(* IEC 61131-3 sources: daoli-st-library/DL_Process (part 10) *)

(* ---- FC_DL_CathodeMillThroughputCalc.st ---- *)
(*
  Component : FC_DL_CathodeMillThroughputCalc
  Category  : DL_Process
  Function  : 粉碎分级产能估算 t/h：由分级轮转速与风量折算，含转速修正与上限钳位
  Complexity: C2
  开源溯源 : DLF 内部原创（R94 族模板派生）；参考语义来源见 SOURCE_HUNTING_MATRIX.md
  规则遵从 : R1-R16
  契约     : 输入 rAirFlowM3h 系统风量 [m3/h]、rSolidsGm3 气流含尘浓度 [g/m3]、
             nWheelRpm 分级轮实际转速 [r/min]、nWheelRefRpm 分级轮额定转速 [r/min]、
             rSpeedExp 转速修正指数 [-]、rCapMaxTh 产能硬上限 [t/h]；
             输出 rThroughputTh 估算产能 [t/h]、rSpeedFactor 转速修正因子 [-]、
             xCapped 触上限、xValid 有效标志、nFaultCode 故障码。
  边界     : 基础产能 = 风量 × 含尘浓度 / 1.0E6（g→t 与 m3/h→t/h 一次换算）；转速因子 =
             (实际/额定)^指数，指数须 >0 且 ≤2；额定转速为分母须 >1.0E-9 [r/min]；
             产能硬限上限必须具备「极限值→REAL 可表性」反算：上限 1.0E4 [t/h] 远小于 REAL 上限 3.4E38，可表。
  码位     : 9801 输入非有限（故障级）；9802 额定转速或指数越域（故障级）。
*)
FUNCTION FC_DL_CathodeMillThroughputCalc : BOOL
VAR_INPUT
    rAirFlowM3h   : LREAL := 5000.0;   // 系统风量 [m3/h] EN: the air volumetric flow of the classifying system
    rSolidsGm3    : LREAL := 200.0;    // 气流含尘浓度 [g/m3] EN: the solids concentration carried by the air
    nWheelRpm     : INT := 3000;       // 分级轮实际转速 [r/min] EN: the actual rotational speed of the classifying wheel
    nWheelRefRpm  : INT := 3000;       // 分级轮额定转速 [r/min] EN: the rated rotational speed of the classifying wheel
    rSpeedExp     : LREAL := 1.0;      // 转速修正指数 [-] EN: the exponent of the speed correction
    rCapMaxTh     : LREAL := 5.0;      // 产能硬上限 [t/h] EN: the hard upper bound of the throughput
END_VAR
VAR_OUTPUT
    rThroughputTh : LREAL;             // 估算产能 [t/h] EN: the estimated throughput in tonnes per hour
    rSpeedFactor  : LREAL;             // 转速修正因子 [-] EN: the speed correction factor
    xCapped       : BOOL;              // 触产能硬上限 EN: the throughput reached the hard upper bound
    xValid        : BOOL;              // 输出可信标志 EN: the outputs are valid
    nFaultCode    : INT;               // 0=无故障 9801=输入非有限 9802=额定转速或指数越域 EN: zero none, 9801 non finite input, 9802 rated speed or exponent out of range
END_VAR
VAR
    xFinAll : BOOL;                    // 浮点入参同时有限 EN: the floating inputs are finite
    rBase   : LREAL;                   // 基础产能（未修正） [t/h] EN: the base throughput before the correction
    rRatio  : LREAL;                   // 转速比 [-] EN: the speed ratio
    rFactor : LREAL;                   // 修正因子中间值 [-] EN: the interim correction factor
    rOut    : LREAL;                   // 产能中间值 [t/h] EN: the interim throughput
END_VAR
VAR CONSTANT
    DL_CMT_Z       : LREAL := 0.0;      // 浮点零常量 EN: the floating point zero constant
    DL_CMT_MILLION : LREAL := 1.0E6;    // 克转吨与每小时一次换算系数 EN: the gram to tonne conversion factor
    DL_CMT_EXP_MAX : LREAL := 2.0;      // 修正指数上限 [-] EN: the upper bound of the exponent
    DL_CMT_MIN     : LREAL := 1.0E-9;   // 分母绝对值下限 EN: the lower bound of the divisor magnitude
    DL_CMT_C_BAD   : INT := 9801;       // 输入非有限 EN: a non finite input
    DL_CMT_C_RANGE : INT := 9802;       // 额定转速或指数越域 EN: the rated speed or the exponent is out of range
END_VAR

// 段1｜出口预置
FC_DL_CathodeMillThroughputCalc := FALSE;   // 返回值预置假 EN: preset the return value to false
rThroughputTh := DL_CMT_Z;                  // 产能预置零 [t/h] EN: preset the throughput to zero
rSpeedFactor := DL_CMT_Z;                   // 修正因子预置零 [-] EN: preset the correction factor to zero
xCapped := FALSE;                           // 触限标志预置假 EN: preset the capped flag to false
xValid := FALSE;                            // 有效标志预置假 EN: preset the validity flag to false
nFaultCode := 0;                            // 故障码预置零 EN: preset the fault code to zero

// 段2｜非有限闸：浮点入参全列（硬上限参与钳位，漏则钳位失效）
xFinAll := (rAirFlowM3h = rAirFlowM3h) AND ((rAirFlowM3h - rAirFlowM3h) = DL_CMT_Z)
        AND (rSolidsGm3 = rSolidsGm3) AND ((rSolidsGm3 - rSolidsGm3) = DL_CMT_Z)
        AND (rSpeedExp = rSpeedExp) AND ((rSpeedExp - rSpeedExp) = DL_CMT_Z)
        AND (rCapMaxTh = rCapMaxTh) AND ((rCapMaxTh - rCapMaxTh) = DL_CMT_Z);   // 四浮点输入有限性 EN: the finiteness of the four floating inputs
IF NOT xFinAll THEN                                                             // 非有限出口 EN: leave early on a non finite input
    nFaultCode := DL_CMT_C_BAD;                                                 // 非有限码 EN: the non finite code
    RETURN;                                                                     // 早退 EN: return early
END_IF

// 段3｜域闸：风量与含尘浓度非负、转速非负、额定转速过分母下限、指数在 (0,2]、硬上限为正
IF (rAirFlowM3h < DL_CMT_Z) OR (rSolidsGm3 < DL_CMT_Z) OR (nWheelRpm < 0) OR (nWheelRefRpm < 0)
   OR (rSpeedExp <= DL_CMT_Z) OR (rSpeedExp > DL_CMT_EXP_MAX) OR (rCapMaxTh <= DL_CMT_Z)
   OR (ABS(INT_TO_LREAL(nWheelRefRpm)) < DL_CMT_MIN) THEN
    nFaultCode := DL_CMT_C_RANGE;                                               // 越域码 EN: the out of range code
    RETURN;                                                                     // 早退 EN: return early
END_IF

// 段4｜主体：基础产能 = 风量 × 含尘 / 1.0E6；因子 = (实际/额定)^指数
rBase := (rAirFlowM3h * rSolidsGm3) / DL_CMT_MILLION;                           // 基础产能 [t/h] EN: the base throughput
rRatio := INT_TO_LREAL(nWheelRpm) / INT_TO_LREAL(nWheelRefRpm);                 // 转速比，分母已证正 [-] EN: the speed ratio, the divisor is proven positive
rFactor := EXP(rSpeedExp * LN(rRatio));                                         // 指数修正 = e^(k·ln r) [-]，避免依赖 EXPT 方言 EN: the exponential correction without a vendor power operator
rOut := rBase * rFactor;                                                        // 修正后产能 [t/h] EN: the corrected throughput

// 段5｜结果复检 + 硬上限钳位（只防上溢，不下抬）
IF (rOut <> rOut) OR (rOut < DL_CMT_Z) THEN                                     // 复检：非有限或负 EN: recheck for a non finite or negative result
    nFaultCode := DL_CMT_C_RANGE;                                               // 复检失败码 EN: the recheck failure code
    RETURN;                                                                     // 早退，出口保持零哨兵 EN: return early with the zero sentinels
END_IF
IF rOut > rCapMaxTh THEN                                                        // 硬上限钳位 EN: the hard upper bound
    rOut := rCapMaxTh;                                                          // 钳到上限 [t/h] EN: clamp to the upper bound
    xCapped := TRUE;                                                            // 置触限标志 EN: raise the capped flag
END_IF

// 段6｜出口
rThroughputTh := rOut;                                                          // 产能出口 [t/h] EN: the throughput output
rSpeedFactor := rFactor;                                                        // 因子出口 [-] EN: the factor output
xValid := TRUE;                                                                 // 结果可信 EN: the results are valid
FC_DL_CathodeMillThroughputCalc := TRUE;                                        // 返回真 EN: return true
END_FUNCTION

(* ---- FC_DL_CathodeMoistureSpecCalc.st ---- *)
(*
  Component : FC_DL_CathodeMoistureSpecCalc
  Category  : DL_Process
  Function  : 水分限值与所需干燥时间反算（一阶指数干燥模型 t = -τ × LN(M目标/M初始)）
  Complexity: C2
  开源溯源 : DLF 内部原创（R94 族模板派生）；参考语义来源见 SOURCE_HUNTING_MATRIX.md
  规则遵从 : R1-R16
  契约     : 输入 rMoistInitPct 初始水分 [%]、rMoistTargetPct 目标水分限值 [%]、
             rDryTauMin 干燥时间常数 [min]、rDryTimeMaxMin 工艺允许最长干燥时间 [min]；
             输出 rDryMin 计算所需干燥时间 [min]、rMoistRatio 水分比 [-]、
             xSpecAchievable 目标在当前允许时间内可达、xValid 有效标志、nFaultCode 故障码。
  边界     : 须 初始水分 > 目标水分 > 0；时间常数为分母须 >1.0E-9 [min]；允许时长须 >0；
             模型不含恒速段与临界含水率，仅适用于降速干燥段（物料表面已不饱和）；
             目标不可达只置 xSpecAchievable=FALSE 为信息级，不置故障。
  码位     : 9801 输入非有限（故障级）；9802 水分关系非法（故障级）；9803 时间常数或允许时长越域（故障级）。
*)
FUNCTION FC_DL_CathodeMoistureSpecCalc : BOOL
VAR_INPUT
    rMoistInitPct   : LREAL := 5.0;      // 初始水分 [%] EN: the initial moisture content
    rMoistTargetPct : LREAL := 0.05;     // 目标水分限值 [%] EN: the target moisture limit
    rDryTauMin      : LREAL := 20.0;     // 干燥时间常数 [min] EN: the drying time constant
    rDryTimeMaxMin  : LREAL := 180.0;    // 工艺允许最长干燥时间 [min] EN: the longest drying time allowed by the process
END_VAR
VAR_OUTPUT
    rDryMin         : LREAL;             // 计算所需干燥时间 [min] EN: the computed drying time required
    rMoistRatio     : LREAL;             // 目标与初始水分之比 [-] EN: the ratio of the target to the initial moisture
    xSpecAchievable : BOOL;              // 目标在允许时间内可达（信息级） EN: the target is reachable within the allowed time, information class only
    xValid          : BOOL;              // 输出可信标志 EN: the outputs are valid
    nFaultCode      : INT;               // 0=无故障 9801=输入非有限 9802=水分关系非法 9803=常数或时长越域 EN: zero none, 9801 non finite, 9802 illegal moisture relation, 9803 constant or duration out of range
END_VAR
VAR
    xFinAll : BOOL;                      // 四输入同时有限 EN: all four inputs are finite
    rRat    : LREAL;                     // 水分比中间值 [-] EN: the interim moisture ratio
    rLn     : LREAL;                     // 水分比对数 [-] EN: the logarithm of the moisture ratio
    rT      : LREAL;                     // 干燥时间中间值 [min] EN: the interim drying time
END_VAR
VAR CONSTANT
    DL_CMS_Z      : LREAL := 0.0;        // 浮点零常量 EN: the floating point zero constant
    DL_CMS_MIN    : LREAL := 1.0E-9;     // 分母绝对值下限 EN: the lower bound of the divisor magnitude
    DL_CMS_C_BAD  : INT := 9801;         // 输入非有限 EN: a non finite input
    DL_CMS_C_REL  : INT := 9802;         // 水分关系非法 EN: an illegal moisture relation
    DL_CMS_C_RANG : INT := 9803;         // 时间常数或允许时长越域 EN: the constant or the duration is out of range
END_VAR

// 段1｜出口预置
FC_DL_CathodeMoistureSpecCalc := FALSE;   // 返回值预置假 EN: preset the return value to false
rDryMin := DL_CMS_Z;                      // 干燥时间预置零 [min] EN: preset the drying time to zero
rMoistRatio := DL_CMS_Z;                  // 水分比预置零 [-] EN: preset the moisture ratio to zero
xSpecAchievable := FALSE;                 // 可达标志预置假 EN: preset the reachability flag to false
xValid := FALSE;                          // 有效标志预置假 EN: preset the validity flag to false
nFaultCode := 0;                          // 故障码预置零 EN: preset the fault code to zero

// 段2｜非有限闸：四输入全列
xFinAll := (rMoistInitPct = rMoistInitPct) AND ((rMoistInitPct - rMoistInitPct) = DL_CMS_Z)
        AND (rMoistTargetPct = rMoistTargetPct) AND ((rMoistTargetPct - rMoistTargetPct) = DL_CMS_Z)
        AND (rDryTauMin = rDryTauMin) AND ((rDryTauMin - rDryTauMin) = DL_CMS_Z)
        AND (rDryTimeMaxMin = rDryTimeMaxMin) AND ((rDryTimeMaxMin - rDryTimeMaxMin) = DL_CMS_Z);   // 四输入有限性 EN: the finiteness of all four inputs
IF NOT xFinAll THEN                                                                                 // 非有限出口 EN: leave early on a non finite input
    nFaultCode := DL_CMS_C_BAD;                                                                     // 非有限码 EN: the non finite code
    RETURN;                                                                                         // 早退 EN: return early
END_IF

// 段3｜域闸：水分关系 初始 > 目标 > 0；时间常数与允许时长为正
IF (rMoistTargetPct <= DL_CMS_Z) OR (rMoistInitPct <= rMoistTargetPct) THEN                          // 水分关系闸 EN: the moisture relation gate
    nFaultCode := DL_CMS_C_REL;                                                                     // 关系非法码 EN: the relation code
    RETURN;                                                                                         // 早退 EN: return early
END_IF
IF (rDryTauMin < DL_CMS_MIN) OR (rDryTimeMaxMin <= DL_CMS_Z) THEN                                    // 常数与时长闸 EN: the constant and duration gate
    nFaultCode := DL_CMS_C_RANG;                                                                    // 越域码 EN: the out of range code
    RETURN;                                                                                         // 早退 EN: return early
END_IF

// 段4｜主体：t = -τ × LN(目标/初始)，比值已证在 (0,1)
rRat := rMoistTargetPct / rMoistInitPct;                                                            // 水分比 [-] EN: the moisture ratio
rLn := LN(rRat);                                                                                    // 水分比对数，已证 <0 [-] EN: the logarithm of the ratio, proven negative
rT := -rDryTauMin * rLn;                                                                            // 所需干燥时间 [min] EN: the drying time required
IF (rT <> rT) OR (rT < DL_CMS_Z) THEN                                                               // 结果复检 EN: recheck the result
    nFaultCode := DL_CMS_C_RANG;                                                                    // 复检失败码 EN: the recheck failure code
    RETURN;                                                                                         // 早退，出口保持零哨兵 EN: return early with the zero sentinels
END_IF

// 段5｜出口：可达性为信息级判据
rDryMin := rT;                                                                                      // 干燥时间出口 [min] EN: the drying time output
rMoistRatio := rRat;                                                                                // 水分比出口 [-] EN: the moisture ratio output
xSpecAchievable := rT <= rDryTimeMaxMin;                                                            // 可达性判定 EN: the reachability verdict
xValid := TRUE;                                                                                     // 结果可信 EN: the results are valid
FC_DL_CathodeMoistureSpecCalc := TRUE;                                                              // 返回真 EN: return true
END_FUNCTION

(* ---- FC_DL_CathodeO2PartialPressureCalc.st ---- *)
(*
  Component : FC_DL_CathodeO2PartialPressureCalc
  Category  : DL_Process
  Function  : 烧结气氛氧分压 = 氧体积浓度 × 总压，并统一换算到 kPa
  Complexity: C2
  开源溯源 : DLF 内部原创（R94 族模板派生）；参考语义来源见 SOURCE_HUNTING_MATRIX.md
  规则遵从 : R1-R16
  契约     : 输入 rO2Pct 氧体积浓度 [%]、rTotalPressKpa 炉膛总压 [kPa]、rO2LowKpa 氧分压下限 [kPa]；
             输出 rPO2Kpa 氧分压 [kPa]、rO2Ppm 氧体积浓度折算 [ppm]、xO2Low 低于下限（信息级）、
             xValid 有效标志、nFaultCode 故障码。
  边界     : 氧浓度须在 0~100 [%] 内、总压须 >std 0（表压与绝压口径由调用方统一为绝压）；
             浓度 1 [%] = 10000 [ppm]，故 ppm = % × 10000；本件为绝压口径，不做大气压叠加。
  码位     : 9801 输入非有限（故障级）；9802 浓度或总压越域（故障级）。
*)
FUNCTION FC_DL_CathodeO2PartialPressureCalc : BOOL
VAR_INPUT
    rO2Pct       : LREAL := 21.0;     // 氧体积浓度 [%] EN: the oxygen volumetric concentration in percent
    rTotalPressKpa: LREAL := 101.325; // 炉膛总压（绝压口径） [kPa] EN: the furnace total pressure on the absolute scale
    rO2LowKpa    : LREAL := 0.5;      // 氧分压工艺下限 [kPa] EN: the technological lower bound of the oxygen partial pressure
END_VAR
VAR_OUTPUT
    rPO2Kpa : LREAL;                  // 氧分压 [kPa] EN: the oxygen partial pressure
    rO2Ppm  : LREAL;                  // 氧体积浓度折算值 [ppm] EN: the oxygen concentration expressed in ppm
    xO2Low  : BOOL;                   // 氧分压低于工艺下限（信息级） EN: the oxygen partial pressure is below the limit, information class only
    xValid  : BOOL;                   // 输出可信标志 EN: the outputs are valid
    nFaultCode : INT;                 // 0=无故障 9801=输入非有限 9802=浓度或总压越域 EN: zero none, 9801 non finite input, 9802 concentration or pressure out of range
END_VAR
VAR
    xFinAll : BOOL;                   // 三输入同时有限 EN: all three inputs are finite
    rFrac   : LREAL;                  // 氧体积分数 [-] EN: the oxygen volumetric fraction
    rPO2    : LREAL;                  // 氧分压中间值 [kPa] EN: the interim oxygen partial pressure
    rPpm    : LREAL;                  // ppm 中间值 [ppm] EN: the interim ppm value
END_VAR
VAR CONSTANT
    DL_COP_Z         : LREAL := 0.0;      // 浮点零常量 EN: the floating point zero constant
    DL_COP_HUNDRED   : LREAL := 100.0;    // 百分数换算系数 EN: the percent conversion factor
    DL_COP_PPM_FACT  : LREAL := 10000.0;  // 百分数转 ppm 的系数 EN: the percent to ppm factor
    DL_COP_C_BAD     : INT := 9801;       // 输入非有限 EN: a non finite input
    DL_COP_C_RANGE   : INT := 9802;       // 浓度或总压越域 EN: the concentration or the pressure is out of range
END_VAR

// 段1｜出口预置
FC_DL_CathodeO2PartialPressureCalc := FALSE;   // 返回值预置假 EN: preset the return value to false
rPO2Kpa := DL_COP_Z;                           // 氧分压预置零 [kPa] EN: preset the partial pressure to zero
rO2Ppm := DL_COP_Z;                            // ppm 预置零 [ppm] EN: preset the ppm value to zero
xO2Low := FALSE;                               // 低压标志预置假 EN: preset the low pressure flag to false
xValid := FALSE;                               // 有效标志预置假 EN: preset the validity flag to false
nFaultCode := 0;                               // 故障码预置零 EN: preset the fault code to zero

// 段2｜非有限闸：三输入全列（下限参与出口判据）
xFinAll := (rO2Pct = rO2Pct) AND ((rO2Pct - rO2Pct) = DL_COP_Z)
        AND (rTotalPressKpa = rTotalPressKpa) AND ((rTotalPressKpa - rTotalPressKpa) = DL_COP_Z)
        AND (rO2LowKpa = rO2LowKpa) AND ((rO2LowKpa - rO2LowKpa) = DL_COP_Z);   // 三输入有限性 EN: the finiteness of all three inputs
IF NOT xFinAll THEN                                                             // 非有限出口 EN: leave early on a non finite input
    nFaultCode := DL_COP_C_BAD;                                                 // 输入非有限码 EN: the non finite code
    RETURN;                                                                     // 早退 EN: return early
END_IF

// 段3｜域闸：氧浓度 0~100 [%]、总压为正、下限非负
IF (rO2Pct < DL_COP_Z) OR (rO2Pct > DL_COP_HUNDRED) OR (rTotalPressKpa <= DL_COP_Z)
   OR (rO2LowKpa < DL_COP_Z) THEN
    nFaultCode := DL_COP_C_RANGE;                                               // 越域码 EN: the out of range code
    RETURN;                                                                     // 早退 EN: return early
END_IF

// 段4｜主体：pO2 = 浓度/100 × 总压；ppm = 浓度 × 10000
rFrac := rO2Pct / DL_COP_HUNDRED;                                               // 氧体积分数 [-] EN: the oxygen volumetric fraction
rPO2 := rFrac * rTotalPressKpa;                                                 // 氧分压 [kPa] EN: the oxygen partial pressure
rPpm := rO2Pct * DL_COP_PPM_FACT;                                               // 浓度转 ppm [ppm] EN: the concentration in ppm

// 段5｜出口
rPO2Kpa := rPO2;                                                                // 氧分压出口 [kPa] EN: the partial pressure output
rO2Ppm := rPpm;                                                                 // ppm 出口 [ppm] EN: the ppm output
xO2Low := rPO2 < rO2LowKpa;                                                     // 低压判据（信息级） EN: the low pressure test, information class only
xValid := TRUE;                                                                 // 结果可信 EN: the results are valid
FC_DL_CathodeO2PartialPressureCalc := TRUE;                                     // 返回真 EN: return true
END_FUNCTION

(* ---- FC_DL_CathodeSaggerLoadCalc.st ---- *)
(*
  Component : FC_DL_CathodeSaggerLoadCalc
  Category  : DL_Process
  Function  : 匣钵装载量 = 层数 × 每层片数 × 单重，并做超重告警
  Complexity: C2
  开源溯源 : DLF 内部原创（R94 族模板派生）；参考语义来源见 SOURCE_HUNTING_MATRIX.md
  规则遵从 : R1-R16
  契约     : 输入 nLayers 层数 [层]、nPerLayer 每层片数 [片/层]、rPieceKg 单片重量 [kg]、
             rMaxLoadKg 匣钵允许装载上限 [kg]；输出 nPieceCount 总片数 [片]、rLoadKg 装载总重 [kg]、
             xOverload 超重（故障级：超重会导致匣钵破裂并损坏辊棒，按安全侧立即判故障）、
             xValid 有效标志、nFaultCode 故障码。
  边界     : 层数与每层片数须在 0~999 内（超过 999 属组态错误，防整数乘法溢出判 9802）；
             单片重量须 ≥0；上限须 >0；总片数 = 层数 × 每层片数，最大 999×999 = 998001 片，INT 可表；
             超重按方向明确判「超上限」，故为故障级（R146：与安全侧一致的异常立即终止）。
  码位     : 9801 输入非有限或为负（故障级）；9802 计数越界（故障级）；9803 超重（故障级）。
*)
FUNCTION FC_DL_CathodeSaggerLoadCalc : BOOL
VAR_INPUT
    nLayers    : INT := 8;           // 匣钵叠放层数 [层] EN: the number of stacked layers in the sagger
    nPerLayer  : INT := 6;           // 每层片数 [片/层] EN: the number of pieces per layer
    rPieceKg   : LREAL := 0.5;       // 单片重量 [kg] EN: the weight of one piece
    rMaxLoadKg : LREAL := 30.0;      // 匣钵允许装载上限 [kg] EN: the allowed load limit of the sagger
END_VAR
VAR_OUTPUT
    nPieceCount : INT;               // 总片数 [片] EN: the total piece count
    rLoadKg     : LREAL;             // 装载总重 [kg] EN: the total load weight
    xOverload   : BOOL;              // 超重（故障级） EN: the load exceeds the limit, a fault class condition
    xValid      : BOOL;              // 输出可信标志 EN: the outputs are valid
    nFaultCode  : INT;               // 0=无故障 9801=输入非法 9802=计数越界 9803=超重 EN: zero none, 9801 illegal input, 9802 count out of range, 9803 overload
END_VAR
VAR
    xFinAll  : BOOL;                 // 两个浮点入参有限 EN: both floating inputs are finite
    nCnt     : INT;                  // 总片数中间值 [片] EN: the interim piece count
    rLoad    : LREAL;                // 总重中间值 [kg] EN: the interim load weight
END_VAR
VAR CONSTANT
    DL_CSL_Z      : LREAL := 0.0;    // 浮点零常量 EN: the floating point zero constant
    DL_CSL_CNT_MAX: INT := 999;      // 层数与每层片数上限 [个] EN: the upper bound of the layer count and the per layer count
    DL_CSL_C_BAD  : INT := 9801;     // 输入非法 EN: an illegal input
    DL_CSL_C_CNT  : INT := 9802;     // 计数越界 EN: the count is out of range
    DL_CSL_C_OVER : INT := 9803;     // 超重 EN: the overload condition
END_VAR

// 段1｜出口预置
FC_DL_CathodeSaggerLoadCalc := FALSE;   // 返回值预置假 EN: preset the return value to false
nPieceCount := 0;                        // 总片数预置零 [片] EN: preset the piece count to zero
rLoadKg := DL_CSL_Z;                     // 总重预置零 [kg] EN: preset the load weight to zero
xOverload := FALSE;                      // 超重标志预置假 EN: preset the overload flag to false
xValid := FALSE;                         // 有效标志预置假 EN: preset the validity flag to false
nFaultCode := 0;                         // 故障码预置零 EN: preset the fault code to zero

// 段2｜非有限闸：两个浮点入参全列（上限参与超重判据）
xFinAll := (rPieceKg = rPieceKg) AND ((rPieceKg - rPieceKg) = DL_CSL_Z)
        AND (rMaxLoadKg = rMaxLoadKg) AND ((rMaxLoadKg - rMaxLoadKg) = DL_CSL_Z);   // 两输入有限性 EN: the finiteness of both inputs
IF NOT xFinAll THEN                                                                 // 非有限出口 EN: leave early on a non finite input
    nFaultCode := DL_CSL_C_BAD;                                                     // 输入非法码 EN: the illegal input code
    RETURN;                                                                         // 早退 EN: return early
END_IF

// 段3｜域闸：单片重量与上限为正、两计数非负且不超 999
IF (rPieceKg < DL_CSL_Z) OR (rMaxLoadKg <= DL_CSL_Z) THEN                            // 数值域闸 EN: the numeric domain gate
    nFaultCode := DL_CSL_C_BAD;                                                     // 输入非法码 EN: the illegal input code
    RETURN;                                                                         // 早退 EN: return early
END_IF
IF (nLayers < 0) OR (nLayers > DL_CSL_CNT_MAX) OR (nPerLayer < 0) OR (nPerLayer > DL_CSL_CNT_MAX) THEN
    nFaultCode := DL_CSL_C_CNT;                                                     // 计数越界码 EN: the count out of range code
    RETURN;                                                                         // 早退 EN: return early
END_IF

// 段4｜主体：片数用整数乘（取值范围已证），重量用标准转换后相乘
nCnt := nLayers * nPerLayer;                                                        // 总片数 [片] EN: the total piece count
rLoad := INT_TO_LREAL(nCnt) * rPieceKg;                                             // 总重 [kg] EN: the total load weight

// 段5｜出口：超重为故障级（安全侧一致的方向明确异常立即终止）
nPieceCount := nCnt;                                                                // 总片数出口 [片] EN: the piece count output
rLoadKg := rLoad;                                                                   // 总重出口 [kg] EN: the load weight output
IF rLoad > rMaxLoadKg THEN                                                          // 超重判据 EN: the overload test
    xOverload := TRUE;                                                              // 置超重标志 EN: raise the overload flag
    nFaultCode := DL_CSL_C_OVER;                                                    // 超重码 EN: the overload code
    xValid := FALSE;                                                                // 超重时输出不可用于投料 EN: the outputs are not usable for loading
    RETURN;                                                                         // 早退（返回假） EN: return false
END_IF
xValid := TRUE;                                                                     // 结果可信 EN: the results are valid
FC_DL_CathodeSaggerLoadCalc := TRUE;                                                // 返回真 EN: return true
END_FUNCTION

(* ---- FC_DL_CathodeSinterSoakCalc.st ---- *)
(*
  Component : FC_DL_CathodeSinterSoakCalc
  Category  : DL_Process
  Function  : 烧结保温时间由固相扩散长度与粒径反算，t = L² / (4D)，含最小值保护
  Complexity: C2
  开源溯源 : DLF 内部原创（R94 族模板派生）；参考语义来源见 SOURCE_HUNTING_MATRIX.md
  规则遵从 : R1-R16
  契约     : 输入 rDiffLenUm 目标扩散长度 [μm]、rDiffCoefUm2Min 有效扩散系数 [μm2/min]、
             rParticleD50Um 一次粒径中位径 [μm]、rSoakMinMin 保温时间下限 [min]；
             输出 rSoakCalcMin 模型计算保温时间 [min]、rSoakMin 施加下限保护后的保温时间 [min]、
             xMinApplied 触底保护生效、xValid 有效标志、nFaultCode 故障码。
  边界     : 扩散系数为分母须 >1.0E-9 [μm2/min]；扩散长度与粒径须 >0；模型 t = L²/(4D)；
             粒径小于两倍扩散长度时扩散已贯穿颗粒，模型外推无意义，rSoakMin 仍给出但不置 xValid=FALSE，
             改由 xMinApplied 与告警表达（本件不设粒径下限门限，交由上层工艺判定）。
  码位     : 9801 输入非法（故障级）；9802 扩散系数过小（故障级）。
*)
FUNCTION FC_DL_CathodeSinterSoakCalc : BOOL
VAR_INPUT
    rDiffLenUm      : LREAL := 2.0;      // 目标固相扩散长度 [μm] EN: the target solid state diffusion length
    rDiffCoefUm2Min : LREAL := 0.05;     // 有效扩散系数 [μm2/min] EN: the effective diffusion coefficient
    rParticleD50Um  : LREAL := 5.0;      // 一次粒径中位径 D50 [μm] EN: the median primary particle size
    rSoakMinMin     : LREAL := 120.0;    // 保温时间工艺下限 [min] EN: the technological lower bound of the soak time
END_VAR
VAR_OUTPUT
    rSoakCalcMin : LREAL;                // 模型计算保温时间 [min] EN: the model computed soak time
    rSoakMin     : LREAL;                // 施加下限保护后的保温时间 [min] EN: the soak time after the lower bound protection
    xMinApplied  : BOOL;                 // 触底保护生效 EN: the lower bound protection took effect
    xThrough     : BOOL;                 // 扩散已贯穿颗粒（信息级） EN: the diffusion length already spans the particle, information class only
    xValid       : BOOL;                 // 输出可信标志 EN: the outputs are valid
    nFaultCode   : INT;                  // 0=无故障 9801=输入非法 9802=扩散系数过小 EN: zero none, 9801 illegal input, 9802 diffusion coefficient too small
END_VAR
VAR
    xFinAll  : BOOL;                     // 四输入同时有限 EN: all four inputs are finite
    rDen     : LREAL;                    // 分母 4D [μm2/min] EN: the divisor, four times the diffusion coefficient
    rSq      : LREAL;                    // 扩散长度平方 [μm2] EN: the squared diffusion length
    rCalc    : LREAL;                    // 计算保温时间 [min] EN: the computed soak time
    rApply   : LREAL;                    // 施加下限后的保温时间 [min] EN: the soak time after the lower bound
END_VAR
VAR CONSTANT
    DL_CSS_Z       : LREAL := 0.0;       // 浮点零常量 EN: the floating point zero constant
    DL_CSS_FOUR    : LREAL := 4.0;       // 扩散方程几何系数 EN: the geometric factor of the diffusion equation
    DL_CSS_TWO     : LREAL := 2.0;       // 贯穿判据倍数 EN: the spanning criterion multiplier
    DL_CSS_MIN     : LREAL := 1.0E-9;    // 分母绝对值下限 [μm2/min] EN: the lower bound of the divisor magnitude
    DL_CSS_C_BAD   : INT := 9801;        // 输入非法 EN: an illegal input
    DL_CSS_C_COEF  : INT := 9802;        // 扩散系数过小 EN: the diffusion coefficient is too small
END_VAR

// 段1｜出口预置
FC_DL_CathodeSinterSoakCalc := FALSE;   // 返回值预置假 EN: preset the return value to false
rSoakCalcMin := DL_CSS_Z;               // 计算保温时间预置零 [min] EN: preset the computed soak time to zero
rSoakMin := DL_CSS_Z;                   // 施加下限后保温时间预置零 [min] EN: preset the final soak time to zero
xMinApplied := FALSE;                   // 触底标志预置假 EN: preset the lower bound flag to false
xThrough := FALSE;                      // 贯穿标志预置假 EN: preset the spanning flag to false
xValid := FALSE;                        // 有效标志预置假 EN: preset the validity flag to false
nFaultCode := 0;                        // 故障码预置零 EN: preset the fault code to zero

// 段2｜非有限闸：四输入全列
xFinAll := (rDiffLenUm = rDiffLenUm) AND ((rDiffLenUm - rDiffLenUm) = DL_CSS_Z)
        AND (rDiffCoefUm2Min = rDiffCoefUm2Min) AND ((rDiffCoefUm2Min - rDiffCoefUm2Min) = DL_CSS_Z)
        AND (rParticleD50Um = rParticleD50Um) AND ((rParticleD50Um - rParticleD50Um) = DL_CSS_Z)
        AND (rSoakMinMin = rSoakMinMin) AND ((rSoakMinMin - rSoakMinMin) = DL_CSS_Z);   // 四输入有限性 EN: the finiteness of all four inputs
IF NOT xFinAll THEN                                                                      // 非有限出口 EN: leave early on a non finite input
    nFaultCode := DL_CSS_C_BAD;                                                          // 输入非法码 EN: the illegal input code
    RETURN;                                                                              // 早退 EN: return early
END_IF

// 段3｜域闸：扩散长度、粒径为正；扩散系数过分母下限；下限时间非负
rDen := DL_CSS_FOUR * rDiffCoefUm2Min;                                                   // 分母 4D [μm2/min] EN: the divisor, four times the diffusion coefficient
IF (rDiffLenUm <= DL_CSS_Z) OR (rParticleD50Um <= DL_CSS_Z) OR (rSoakMinMin < DL_CSS_Z)
   OR (ABS(rDen) < DL_CSS_MIN) THEN
    nFaultCode := DL_CSS_C_COEF;                                                         // 系数或域非法码 EN: the coefficient or domain code
    RETURN;                                                                              // 早退 EN: return early
END_IF

// 段4｜主体：t = L² / (4D)
rSq := rDiffLenUm * rDiffLenUm;                                                          // 扩散长度平方 [μm2] EN: the squared diffusion length
rCalc := rSq / rDen;                                                                     // 计算保温时间 [min] EN: the computed soak time
IF (rCalc <> rCalc) OR (rCalc < DL_CSS_Z) THEN                                           // 结果复检 EN: recheck the result
    nFaultCode := DL_CSS_C_COEF;                                                         // 复检失败码 EN: the recheck failure code
    RETURN;                                                                              // 早退，出口保持零哨兵 EN: return early with the zero sentinels
END_IF

// 段5｜最小值保护与贯穿标记
rApply := rCalc;                                                                         // 施加下限工作副本 [min] EN: the working copy for the lower bound
xMinApplied := rCalc < rSoakMinMin;                                                      // 触底判据 EN: the lower bound test
IF xMinApplied THEN                                                                      // 触底则抬到工艺下限 EN: raise to the process lower bound
    rApply := rSoakMinMin;                                                               // 施加下限 [min] EN: apply the lower bound
END_IF
xThrough := rDiffLenUm >= (rParticleD50Um / DL_CSS_TWO);                                 // 贯穿判据（信息级） EN: the spanning test, information class only

// 段6｜出口
rSoakCalcMin := rCalc;                                                                   // 计算值出口 [min] EN: the computed value output
rSoakMin := rApply;                                                                      // 最终值出口 [min] EN: the final value output
xValid := TRUE;                                                                          // 结果可信 EN: the results are valid
FC_DL_CathodeSinterSoakCalc := TRUE;                                                     // 返回真 EN: return true
END_FUNCTION

(* ---- FC_DL_CathodeTapDensityCalc.st ---- *)
(*
  Component : FC_DL_CathodeTapDensityCalc
  Category  : DL_Process
  Function  : 振实密度 = 质量 / 振实后体积，并按振次做修正
  Complexity: C2
  开源溯源 : DLF 内部原创（R94 族模板派生）；参考语义来源见 SOURCE_HUNTING_MATRIX.md
  规则遵从 : R1-R16
  契约     : 输入 rMassG 试样质量 [g]、rVolumeMl 振实后体积 [ml]、nTaps 实测振次 [次]、
             nRefTaps 标准振次 [次]、rTapCoef 振次修正系数 [-]；
             输出 rDensityGml 实测振实密度 [g/ml]、rDensityCorrGml 修正到标准振次的密度 [g/ml]、
             xValid 有效标志、nFaultCode 故障码。
  边界     : 体积为分母须 >1.0E-9 [ml]；振次须 ≥1（取对数的前提），标准振次须 ≥1；
             修正模型 rho_ref = rho × (1 + k × LN(nRef/nTaps))，k 须在 [0, 0.2] 内，
             越域判 9803（k 越域会把修正放大成伪数据）；1 g/ml = 1 g/cm3，单位不做换算。
  码位     : 9801 输入非法（故障级）；9802 体积过小或振次非法（故障级）；9803 修正系数越域（故障级）。
*)
FUNCTION FC_DL_CathodeTapDensityCalc : BOOL
VAR_INPUT
    rMassG    : LREAL := 100.0;    // 试样质量 [g] EN: the mass of the sample
    rVolumeMl : LREAL := 50.0;     // 振实后体积 [ml] EN: the tapped volume of the sample
    nTaps     : INT := 3000;       // 实测振次 [次] EN: the tap count actually applied
    nRefTaps  : INT := 3000;       // 标准振次 [次] EN: the reference tap count
    rTapCoef  : LREAL := 0.02;     // 振次修正系数 [-] EN: the tap count correction coefficient
END_VAR
VAR_OUTPUT
    rDensityGml     : LREAL;       // 实测振实密度 [g/ml] EN: the measured tap density
    rDensityCorrGml : LREAL;       // 修正到标准振次的密度 [g/ml] EN: the density corrected to the reference tap count
    xValid          : BOOL;        // 输出可信标志 EN: the outputs are valid
    nFaultCode      : INT;         // 0=无故障 9801=输入非法 9802=体积或振次非法 9803=系数越域 EN: zero none, 9801 illegal input, 9802 volume or taps illegal, 9803 coefficient out of range
END_VAR
VAR
    xFinAll : BOOL;                // 三个浮点入参有限 EN: the three floating inputs are finite
    rDen    : LREAL;               // 分母（振实后体积） [ml] EN: the divisor, the tapped volume
    rRho    : LREAL;               // 实测密度 [g/ml] EN: the measured density
    rLnCorr : LREAL;               // 振次比对数 [-] EN: the logarithm of the tap ratio
    rCorr   : LREAL;               // 密度修正中间值 [g/ml] EN: the interim corrected density
END_VAR
VAR CONSTANT
    DL_CTD_Z        : LREAL := 0.0;   // 浮点零常量 EN: the floating point zero constant
    DL_CTD_ONE      : LREAL := 1.0;   // 浮点壹常量 EN: the floating point one constant
    DL_CTD_COEF_MAX : LREAL := 0.2;   // 修正系数上限 [-] EN: the upper bound of the correction coefficient
    DL_CTD_MIN      : LREAL := 1.0E-9;// 分母绝对值下限 [ml] EN: the lower bound of the divisor magnitude
    DL_CTD_C_BAD    : INT := 9801;    // 输入非法 EN: an illegal input
    DL_CTD_C_DEN    : INT := 9802;    // 体积过小或振次非法 EN: the volume is too small or the taps are illegal
    DL_CTD_C_COEF   : INT := 9803;    // 修正系数越域 EN: the coefficient is out of range
END_VAR

// 段1｜出口预置
FC_DL_CathodeTapDensityCalc := FALSE;   // 返回值预置假 EN: preset the return value to false
rDensityGml := DL_CTD_Z;                 // 实测密度预置零 [g/ml] EN: preset the measured density to zero
rDensityCorrGml := DL_CTD_Z;             // 修正密度预置零 [g/ml] EN: preset the corrected density to zero
xValid := FALSE;                         // 有效标志预置假 EN: preset the validity flag to false
nFaultCode := 0;                         // 故障码预置零 EN: preset the fault code to zero

// 段2｜非有限闸：三浮点入参全列
xFinAll := (rMassG = rMassG) AND ((rMassG - rMassG) = DL_CTD_Z)
        AND (rVolumeMl = rVolumeMl) AND ((rVolumeMl - rVolumeMl) = DL_CTD_Z)
        AND (rTapCoef = rTapCoef) AND ((rTapCoef - rTapCoef) = DL_CTD_Z);   // 三输入有限性 EN: the finiteness of all three inputs
IF NOT xFinAll THEN                                                        // 非有限出口 EN: leave early on a non finite input
    nFaultCode := DL_CTD_C_BAD;                                            // 输入非法码 EN: the illegal input code
    RETURN;                                                                // 早退 EN: return early
END_IF

// 段3｜域闸：质量为非负、体积过分母下限、振次 ≥1
rDen := rVolumeMl;                                                          // 取分母 [ml] EN: take the divisor
IF (rMassG < DL_CTD_Z) OR (ABS(rDen) < DL_CTD_MIN) OR (nTaps < 1) OR (nRefTaps < 1) THEN
    nFaultCode := DL_CTD_C_DEN;                                            // 体积或振次非法码 EN: the volume or tap code
    RETURN;                                                                // 早退 EN: return early
END_IF
IF (rTapCoef < DL_CTD_Z) OR (rTapCoef > DL_CTD_COEF_MAX) THEN               // 系数域闸 EN: the coefficient domain gate
    nFaultCode := DL_CTD_C_COEF;                                            // 系数越域码 EN: the coefficient code
    RETURN;                                                                // 早退 EN: return early
END_IF

// 段4｜主体：实测密度与振次修正（两出口同源，修正只缩放实测值不另起公式）
rRho := rMassG / rDen;                                                      // 实测振实密度 [g/ml] EN: the measured tap density
rLnCorr := LN(INT_TO_LREAL(nRefTaps) / INT_TO_LREAL(nTaps));                // 振次比对数 [-]，两者已证 ≥1 EN: the logarithm of the tap ratio
rCorr := rRho * (DL_CTD_ONE + rTapCoef * rLnCorr);                          // 修正密度 [g/ml] EN: the corrected density
IF (rCorr <> rCorr) OR (rCorr < DL_CTD_Z) THEN                              // 结果复检 EN: recheck the result
    nFaultCode := DL_CTD_C_COEF;                                            // 复检失败码 EN: the recheck failure code
    rDensityGml := rRho;                                                    // 实测值仍可给出 EN: the measured value is still published
    RETURN;                                                                // 早退 EN: return early
END_IF

// 段5｜出口
rDensityGml := rRho;                                                        // 实测密度出口 [g/ml] EN: the measured density output
rDensityCorrGml := rCorr;                                                   // 修正密度出口 [g/ml] EN: the corrected density output
xValid := TRUE;                                                             // 结果可信 EN: the results are valid
FC_DL_CathodeTapDensityCalc := TRUE;                                        // 返回真 EN: return true
END_FUNCTION

(* ---- FC_DL_CellOccupyRateCalc.st ---- *)
(*
  ============================================================
  组件名 : FC_DL_CellOccupyRateCalc
  分类   : DL_Process
  功能   : 货位占用率计算，扣除封存货位后按可用货位求占用百分比与空闲数
  复杂度 : C1
  版本   : 1.0.0
  作者   : 道莅工业代码库工厂 / R81
  日期   : 2026-11-24
  开源溯源 : clean-room（no upstream）—— 依据公开工程公式自研，未复制任何上游实现
  红线自检 : R1 无GVL/R2 无物理地址/R3 纯IEC/R4 防除零/R5 双语注释
  接口说明 :
      可用货位 = 总货位 - 封存货位；占用率 = 已用 / 可用 * 100。
      可用货位 <= 0 时占用率无定义，直接判无效，不输出替代值。
      空闲货位 = 可用 - 已用，小于 0 表示超占（数据异常），本实现按 0 截断并保持比例可算。
      中间量用 DINT 承载，避免 INT 减法溢出。
  ============================================================
*)
FUNCTION FC_DL_CellOccupyRateCalc : BOOL
VAR_INPUT
    bEnable       : BOOL; // 使能：TRUE 时计算 / Enable: TRUE to compute
    bErr          : BOOL; // 外部故障：TRUE 时立即退出并置结果无效 / External fault: TRUE aborts with invalid result
    iCellTotal    : INT;  // 货位总数量 [个] / total number of storage cells [unit]
    iCellUsed     : INT;  // 已占用货位数量 [个] / number of occupied cells [unit]
    iCellBlocked  : INT;  // 封存禁用货位数量 [个] / number of blocked or disabled cells [unit]
END_VAR
VAR_OUTPUT
    rOccupyPct : REAL; // 可用货位占用率 [%] / occupancy rate over the available cells [percent]
    iCellFree  : INT;  // 空闲货位数量，负值按 0 截断 [个] / free cell count, negative clamped to zero [unit]
    iCellAvail : INT;  // 扣除封存后的可用货位数量 [个] / available cell count after removing blocked cells [unit]
    bValid     : BOOL; // 输出有效：TRUE 表示结果可用 / Output valid
END_VAR
VAR CONSTANT
    DL_R_MAX : REAL := 3.0E38;  // 实数上界，用于拦截 Inf [无量纲] / real upper bound used to reject infinity [dimensionless]
    DL_EPS   : REAL := 1.0E-12; // 除零判定阈值 [无量纲] / division guard threshold [dimensionless]
    DL_PCT   : REAL := 100.0;   // 百分数换算系数 [无量纲] / percentage scaling factor [dimensionless]
END_VAR
VAR
    _diAvail : DINT := 0; // 可用货位中间量，DINT 防溢出 [个] / intermediate available count in DINT [unit]
    _diFree  : DINT := 0; // 空闲货位中间量，DINT 防溢出 [个] / intermediate free count in DINT [unit]
    _rAvail  : REAL := 0.0; // 可用货位折算实数 [个] / available count cast to real [unit]
END_VAR

    // 段 1｜出口预置
    rOccupyPct := 0.0;
    iCellFree := 0;
    iCellAvail := 0;
    bValid := FALSE;
    // 段 2｜使能闸与外部故障闸
    IF NOT bEnable THEN
        RETURN;
    END_IF;
    IF bErr THEN
        RETURN;
    END_IF;
    // 段 3｜域闸：总数必须为正，已用与封存不得为负
    IF iCellTotal <= 0 THEN
        RETURN;
    END_IF;
    IF (iCellUsed < 0) OR (iCellBlocked < 0) THEN
        RETURN;
    END_IF;
    // 段 4｜可用货位：总数减封存
    _diAvail := INT_TO_DINT(iCellTotal) - INT_TO_DINT(iCellBlocked);
    // 段 5｜可用货位非正闸：此时占用率无定义，判无效
    IF _diAvail <= 0 THEN
        bValid := FALSE;
        FC_DL_CellOccupyRateCalc := bValid;
        RETURN;
    END_IF;
    iCellAvail := DINT_TO_INT(_diAvail);
    // 段 6｜空闲货位：超占按 0 截断
    _diFree := _diAvail - INT_TO_DINT(iCellUsed);
    IF _diFree < 0 THEN
        _diFree := 0;
    END_IF;
    iCellFree := DINT_TO_INT(_diFree);
    // 段 7｜占用率
    _rAvail := DINT_TO_REAL(_diAvail);
    IF ABS(_rAvail) <= DL_EPS THEN
        RETURN;
    END_IF;
    rOccupyPct := INT_TO_REAL(iCellUsed) / _rAvail * DL_PCT;
    bValid := TRUE;
    FC_DL_CellOccupyRateCalc := bValid;
END_FUNCTION

(* ---- FC_DL_CentrateTurbidityIdx.st ---- *)
(*
  道莅工业代码库 / Daoli Industrial ST Library
  组件: FC_DL_CentrateTurbidityIdx
  分类: DL_Process
  开源溯源: 无（clean-room 工程公式自研；参考公开工艺计算公式，未复制任何受版权保护代码）
  许可证: 本项目自有 (MIT)
  功能: 离心液（分离液）浊度相对基线指数与跑料（携带固体）判定
*)
FUNCTION FC_DL_CentrateTurbidityIdx : BOOL
VAR_INPUT
    rNtuNow : REAL; // 当前离心液浊度 [NTU] / current centrate turbidity
    rNtuBase : REAL; // 清洁运行基线浊度 [NTU] / clean-operation baseline turbidity
    rNtuLimit : REAL; // 跑料报警浊度门槛 [NTU] / carry-over alarm threshold
END_VAR
VAR_OUTPUT
    rIdx : REAL; // 浊度指数 = 当前/基线 [-]，1.0 = 与基线持平 / turbidity index, 1.0 equals baseline
    bValid : BOOL; // 结果有效位 [-] / result valid flag
    bCarryOver : BOOL; // 跑料标志（浊度超门槛）[-] / solids carry-over flag
    iErrCode : INT; // 事件码 0=正常 1=基线浊度非法 2=指数超可观测上限 3=结果非有限 / event code
END_VAR
VAR CONSTANT
    rIdxCap : REAL := 1000.0; // 指数输出饱和上限 [-] / index saturation cap
END_VAR
VAR
    rIdxRaw : REAL; // 未限幅指数 [-] / unlimited index
END_VAR

    // —— 段 0：全路径预清 —— //
    rIdxRaw := 0.0;
    rIdx := 0.0;
    bValid := FALSE;
    bCarryOver := FALSE;
    iErrCode := 0;
    FC_DL_CentrateTurbidityIdx := FALSE;
    // —— 段 1：分母闸（基线浊度，清洗后近零会导致指数爆炸） —— //
    IF rNtuBase <= 0.0 THEN
        iErrCode := 1; // 基线浊度非法，指数无定义 / invalid baseline, index undefined
        RETURN;
    END_IF;
    // —— 段 2：量纲链 (NTU)/(NTU) = 无量纲指数 —— //
    rIdxRaw := rNtuNow / rNtuBase; // 浊度指数 [-] / turbidity index
    // —— 段 3：结果域闸、负值防御与饱和 —— //
    IF ABS(rIdxRaw) > 1.0E15 THEN
        iErrCode := 3; // 结果非有限，强制归零 / non-finite result, forced to zero
        RETURN;
    END_IF;
    IF rIdxRaw < 0.0 THEN
        rIdx := 0.0; // 负浊度不可能，钳零 / negative turbidity impossible
    ELSIF rIdxRaw > rIdxCap THEN
        rIdx := rIdxCap; // 超可观测上限饱和 / saturate at observable cap
        iErrCode := 2; // 信息级：指数超上限，基线可能失效 / info: index capped, baseline suspect
    ELSE
        rIdx := rIdxRaw;
    END_IF;
    // —— 段 4：跑料判定（比较用原始浊度，不用饱和后的指数） —— //
    bCarryOver := rNtuNow > rNtuLimit; // 跑料标志 [-] / carry-over flag
    bValid := TRUE;
    FC_DL_CentrateTurbidityIdx := TRUE;
END_FUNCTION

(* ---- FC_DL_CipCausticStrengthCalc.st ---- *)
// FC_DL_CipCausticStrengthCalc v1.0.0
// 开源溯源：clean-room 自研（族 DL_Process，ST 生态实测 0 命中，无外部代码引入）
(*
  功能: CIP 碱液调配：目标碱量 = 目标浓度·液量/100 [L·%]，当前碱量 = 当前浓度·液量/100，
        缺额 = 目标 − 当前，补浓碱体积 = 缺额/(浓碱浓度 − 目标浓度) [L]（稀释到目标的物料平衡）；
        当前浓度高于目标时补水体积 = 液量·(当前/目标 − 1) [L]。两工况互斥。
  邻件/码位: 与 FC_DL_KegFillingCounterPressureCalc 同属灌装/清洗线设备件（CIP 化学 vs 灌装压力）；
             16#0002_9238 = 非有限、目标浓度越界、液量非正、当前浓度为负或补碱补水互斥违例。
*)
FUNCTION FC_DL_CipCausticStrengthCalc : REAL
VAR_INPUT
    fConcNow    : REAL := 1.5;      // 当前碱液浓度 [%]，域 >= 0 / Current concentration [%]
    fVolNow     : REAL := 2000.0;   // 当前液量 [L]，域 > 0 / Current volume [L]
    fConcTarget : REAL := 2.0;      // 目标浓度 [%]，域 (0, 浓碱浓度) / Target concentration [%]
    fConcStock  : REAL := 30.0;     // 浓碱浓度 [%]，域 > 目标浓度 / Stock concentration [%]
END_VAR
VAR_OUTPUT
    fAddVol   : REAL;               // 需补浓碱体积 [L] / Stock caustic to add [L]
    fAddWater : REAL;               // 需补水体积 [L] / Water to add [L]
    bValid    : BOOL;               // 结果有效回执 [-] / Result validity receipt
    uErrorId  : UDINT;              // 事件码，0 = 无事件 / Event code
END_VAR
VAR
    fAlkaliGap : REAL := 0.0;       // 碱量缺额 [L·%] / Alkali deficit [L percent]
END_VAR
// 段 0：全路径出口安全缺省 / Safe defaults on all outlets
fAddVol := 0.0;                     // 补碱体积缺省零 / Stock caustic default zero
fAddWater := 0.0;                   // 补水体积缺省零 / Water to add default zero
bValid := FALSE;                    // 有效回执预清 / Validity preset clear
uErrorId := 16#0000;                // 事件码预清 / Event code preset clear
FC_DL_CipCausticStrengthCalc := 0.0;    // 返回值缺省零（镜像补碱体积）/ Return default zero
// 段 1：非有限闸（四入参全枚举）/ Non-finite gate over all inputs
IF (fConcNow <> fConcNow) OR (fVolNow <> fVolNow)
   OR (fConcTarget <> fConcTarget) OR (fConcStock <> fConcStock)
   OR (ABS(fConcNow) >= 3.0E38) OR (ABS(fVolNow) >= 3.0E38)
   OR (ABS(fConcTarget) >= 3.0E38) OR (ABS(fConcStock) >= 3.0E38) THEN
    uErrorId := 16#0002_9238;   // 入参非有限拒收 / Non-finite input reject
    RETURN;
END_IF
// 段 2：域闸（目标浓度区间 + 液量正 + 当前浓度非负，R4）/ Domain gate
IF (fConcTarget <= 1.0E-6) OR (fConcTarget >= fConcStock) THEN
    uErrorId := 16#0002_9238;   // 目标浓度越界（分母近零）/ Target concentration out of range
    RETURN;
END_IF
IF fVolNow <= 1.0E-6 THEN
    uErrorId := 16#0002_9238;   // 液量非正 / Non-positive liquid volume
    RETURN;
END_IF
IF fConcNow < 0.0 THEN
    uErrorId := 16#0002_9238;   // 当前浓度为负 / Negative current concentration
    RETURN;
END_IF
// 段 3：主计算（碱量差 → 补碱体积 / 补水体积，两工况互斥）/ Main computation
// 碱量衡算（R92-修正）：(C_n·V + C_s·x)/(V+x) = C_t  ⇒  x = (C_t − C_n)·V/(C_s − C_t)
// 说明：早期版本误把缺额再除 100（浓度已按 % 计），致补碱量偏小 100 倍、CIP 永久欠配
fAlkaliGap := (fConcTarget - fConcNow) * fVolNow;               // 碱量缺额 [%·L] / Alkali deficit
IF fAlkaliGap > 1.0E-6 THEN
    fAddVol := fAlkaliGap / (fConcStock - fConcTarget);          // 补浓碱体积 [L] / Stock to add
END_IF
IF fConcNow > fConcTarget THEN
    fAddWater := fVolNow * (fConcNow / fConcTarget - 1.0);       // 补水体积 [L] / Water to add
END_IF
// 段 4：出口闸（非有限复核 + 非负复核 + 互斥复核）/ Outlet gate
IF (fAddVol <> fAddVol) OR (fAddWater <> fAddWater)
   OR (ABS(fAddVol) >= 3.0E38) OR (ABS(fAddWater) >= 3.0E38)
   OR (fAddVol < 0.0) OR (fAddWater < 0.0)
   OR ((fAddVol > 1.0E-6) AND (fAddWater > 1.0E-6)) THEN
    fAddVol := 0.0;             // 复核失败回缺省（含互斥违例）/ Fallback on recheck failure
    fAddWater := 0.0;           // 复核失败回缺省（含互斥违例）/ Fallback on recheck failure
    uErrorId := 16#0002_9238;   // 出口复核拒收 / Output recheck reject
    RETURN;
END_IF
bValid := TRUE;                 // 有效回执 / Validity receipt
FC_DL_CipCausticStrengthCalc := fAddVol;        // 返回值镜像补碱体积 / Return mirrors stock volume
END_FUNCTION

(* ---- FC_DL_ClarifierSurfaceLoad.st ---- *)
(*
  道莅工业代码库 / Daoli Industrial ST Library
  组件: FC_DL_ClarifierSurfaceLoad
  分类: DL_Process
  开源溯源: 无（clean-room 工程公式自研；参考公开工艺计算公式，未复制任何受版权保护代码）
  许可证: 本项目自有 (MIT)
  功能: 沉淀池表面水力负荷计算与上限越限判定
*)
FUNCTION FC_DL_ClarifierSurfaceLoad : BOOL
VAR_INPUT
    rFlowM3h : REAL; // 进水流量 [m3/h] / influent flow
    rAreaM2 : REAL; // 沉淀池有效沉淀面积 [m2] / effective settling area
    rLimitM3m2h : REAL; // 表面负荷设计上限 [m3/(m2·h)] / design surface loading limit
END_VAR
VAR_OUTPUT
    rLoadM3m2h : REAL; // 表面水力负荷 [m3/(m2·h)] / surface hydraulic loading
    bValid : BOOL; // 结果有效位 [-] / result valid flag
    bOver : BOOL; // 越限标志（负荷高于设计上限）[-] / over-limit flag
    iErrCode : INT; // 事件码 0=正常 1=面积非法 2=结果非有限 / event code
END_VAR
VAR
    rLoadRaw : REAL; // 未限幅负荷 [m3/(m2·h)] / unlimited loading
END_VAR

    // —— 段 0：全路径预清 —— //
    rLoadRaw := 0.0;
    rLoadM3m2h := 0.0;
    bValid := FALSE;
    bOver := FALSE;
    iErrCode := 0;
    FC_DL_ClarifierSurfaceLoad := FALSE;
    // —— 段 1：分母闸（沉淀面积必须为正） —— //
    IF rAreaM2 <= 0.0 THEN
        iErrCode := 1; // 面积非法，负荷无定义 / invalid area, loading undefined
        RETURN;
    END_IF;
    // —— 段 2：量纲链 (m3/h)/(m2) = m3/(m2·h) —— //
    rLoadRaw := rFlowM3h / rAreaM2; // 表面负荷 [m3/(m2·h)] / surface loading
    // —— 段 3：结果域闸（非有限即归零作废） —— //
    IF ABS(rLoadRaw) > 1.0E15 THEN
        iErrCode := 2; // 结果非有限，强制归零 / non-finite result, forced to zero
        RETURN;
    END_IF;
    // —— 段 4：负流量防御与出参收口 —— //
    IF rLoadRaw < 0.0 THEN
        rLoadM3m2h := 0.0; // 负流量无物理意义 / negative flow is unphysical
    ELSE
        rLoadM3m2h := rLoadRaw;
    END_IF;
    bOver := rLoadM3m2h > rLimitM3m2h; // 越限判定 [-] / over-limit test
    bValid := TRUE;
    FC_DL_ClarifierSurfaceLoad := TRUE;
END_FUNCTION

(* ---- FC_DL_ClinkerCoolingRateCalc.st ---- *)
(*
  Name: FC_DL_ClinkerCoolingRateCalc
  Category: DL_Process
  Version: 1.0.0
  Round: R91 / 2026-11-25
  开源溯源：clean-room 自研（族 水泥窑篦冷机与预热器，ST 开源生态实测 0 命中，无外部代码引入）
  功能：1) 熟料冷却速率按「两测温点温差除以停留时间」计算，单位统一折算为 K/min：
           fRateKmin = (fTempUpC − fTempDownC) / fDwellMin，
           停留时间已在引脚上以分钟给出（min），故无需再乘 60，避免二次折算引入量纲错误。
        2) 速率上下限约束由 fRateLoKmin / fRateHiKmin 给出：低于下限说明冷却不足
           （急冷段不够，C3S 晶型转化不充分、易磨性变差）；高于上限说明冷却过激
           （篦床拉速过快或风量过大，篦板热应力与磨损加剧）。
        3) 输出温差 fDropK 与速率 fRateKmin，两个方向越限位各占一个布尔，便于上层分别处置。
  边界条件：1) 非有限值闸：四路实值入参先过 NOT(x > -DL_BIG AND x < DL_BIG)，同时拦 NaN 与 Inf，
           命中即闸断实值通路（全部输出强制 0.0），不得只置标志（R19）。
        2) 时间零闸：停留时间 fDwellMin <= DL_EPS 时不做除法（分母为零），判无效并清零全部输出。
        3) 温差方向闸：fTempUpC 必须严格高于 fTempDownC，温差为负属测点接反或标签错位，判无效，
           不取绝对值掩盖符号错误（取绝对值会把接反的测点伪装成正常冷却）。
        4) 限值域闸：0.0 <= fRateLoKmin < fRateHiKmin，否则上下限判据同时失效，视为组态错误判无效。
        5) 判据取原始值（R24）：越限判定使用钳制前的 _fRateRawKmin，不得先钳再判。
        6) 物理域钳制：速率钳 0.0 ~ DL_RATE_HI_KMIN；温差钳 >= 0。
  量纲自证：fDropK = (degC) − (degC) = (K)；
           fRateKmin = (K)/(min) = K/min，与 fRateLoKmin / fRateHiKmin 同量纲 [K/min]，可直接比较。
  修订历史 Revision :
    2026-11-25  v1.0.0  R91 首版
*)

FUNCTION FC_DL_ClinkerCoolingRateCalc : BOOL
VAR_INPUT
    fTempUpC         : REAL;   // 上游测点熟料温度 [degC] / Upstream clinker temperature [degC]
    fTempDownC       : REAL;   // 下游测点熟料温度 [degC] / Downstream clinker temperature [degC]
    fDwellMin        : REAL;   // 两测点间熟料停留时间 [min] / Clinker dwell time between the two points [min]
    fRateLoKmin      : REAL;   // 冷却速率工艺下限 [K/min] / Cooling rate process low limit [K/min]
    fRateHiKmin      : REAL;   // 冷却速率工艺上限 [K/min] / Cooling rate process high limit [K/min]
END_VAR
VAR_OUTPUT
    fRateKmin        : REAL;   // 熟料冷却速率 [K/min] / Clinker cooling rate [K/min]
    fDropK           : REAL;   // 两测点温差 [K] / Temperature drop across the two points [K]
    xRateLow         : BOOL;   // 速率低于下限标志 [bool] / Rate below low limit flag [bool]
    xRateHigh        : BOOL;   // 速率高于上限标志 [bool] / Rate above high limit flag [bool]
    xValid           : BOOL;   // 计算有效标志 [bool] / Calculation valid flag [bool]
END_VAR
VAR
    _fDropRawK       : REAL;   // 钳制前的温差 [K] / Raw temperature drop [K]
    _fRateRawKmin    : REAL;   // 钳制前的原始速率 [K/min] / Raw cooling rate before limiting [K/min]
END_VAR
VAR CONSTANT
    DL_EPS           : REAL := 1.0E-9;    // 数值零闸阈值 [-] / Numeric zero gate threshold [-]
    DL_BIG           : REAL := 1.0E12;    // 非有限值闸量级上限 [-] / Finiteness gate magnitude [-]
    DL_MIN_PER_MIN   : REAL := 1.0;       // 分钟基准折算（引脚已为 min）[min/min] / Minute basis, pin already in minutes [min/min]
    DL_RATE_HI_KMIN  : REAL := 500.0;     // 冷却速率物理上限 [K/min] / Cooling rate physical upper bound [K/min]
    DL_ZERO_K        : REAL := 0.0;       // 温差零基准 [K] / Zero temperature-difference reference [K]
END_VAR

(* —— 段 1：非有限值闸（R19：闸断实值通路） —— *)
IF NOT (fTempUpC > -DL_BIG AND fTempUpC < DL_BIG)
   OR NOT (fTempDownC > -DL_BIG AND fTempDownC < DL_BIG)
   OR NOT (fDwellMin > -DL_BIG AND fDwellMin < DL_BIG)
   OR NOT (fRateLoKmin > -DL_BIG AND fRateLoKmin < DL_BIG)
   OR NOT (fRateHiKmin > -DL_BIG AND fRateHiKmin < DL_BIG) THEN
    fRateKmin := 0.0;                       // 输出强制 0.0，切断污染源 / Force zero, cut polluted path
    fDropK := 0.0;                          // 温差强制 0.0 / Drop forced to zero
    xRateLow := FALSE;                      // 失效侧越限位保持假 / Limit flags stay false
    xRateHigh := FALSE;                     // 失效侧越限位保持假 / Limit flags stay false
    xValid := FALSE;                        // 有效位清零 / Validity cleared
    FC_DL_ClinkerCoolingRateCalc := FALSE;  // 返回码与有效位同源 / Return mirrors validity
    RETURN;                                 // 立即退出 / Immediate exit
END_IF

(* —— 段 2：时间零闸与限值域闸（分母为停留时间） —— *)
IF (fDwellMin <= DL_EPS)                                          // 停留时间不可为零
   OR (fRateLoKmin < 0.0)                                         // 下限不得为负
   OR (fRateHiKmin <= fRateLoKmin) THEN                           // 上限必须严格大于下限
    fRateKmin := 0.0;                       // 分母为零即速率不可算 / No dwell, no rate
    fDropK := 0.0;                          // 温差不可用 / Drop not usable
    xRateLow := FALSE;                      // 越限位保持假 / Limit flags stay false
    xRateHigh := FALSE;                     // 越限位保持假 / Limit flags stay false
    xValid := FALSE;                        // 判无效 / Invalid
    FC_DL_ClinkerCoolingRateCalc := FALSE;  // 返回码同步 / Return synchronised
    RETURN;                                 // 提前退出 / Early exit
END_IF

(* —— 段 3：主算式（不钳制，先出原始值供段 4 判据使用，R24） —— *)
_fDropRawK := fTempUpC - fTempDownC;                                              // 两测点温差 [K]
_fRateRawKmin := _fDropRawK / fDwellMin * DL_MIN_PER_MIN;                          // 冷却速率 [K/min]

(* —— 段 4：判据（取原始值；单点 BOOL 聚合避免多处赋 FALSE 覆盖） —— *)
xRateLow := (_fRateRawKmin < fRateLoKmin);                                        // 低于工艺下限
xRateHigh := (_fRateRawKmin > fRateHiKmin);                                       // 高于工艺上限
xValid := (fRateLoKmin >= 0.0)                                                    // 下限须非负（已验）
          AND (fRateHiKmin <= DL_RATE_HI_KMIN)                                    // 上限不得超物理上限
          AND (_fDropRawK > DL_ZERO_K)                                            // 下游必须比上游冷（方向固定）
          AND (_fRateRawKmin >= DL_ZERO_K);                                       // 速率不得为负

(* —— 段 5：输出单点写盘（钳制到物理域内，判定结果已在段 4 定案） —— *)
fRateKmin := LIMIT(0.0, _fRateRawKmin, DL_RATE_HI_KMIN);                           // 速率钳 0..物理上限 [K/min]
fDropK := MAX(DL_ZERO_K, _fDropRawK);                                              // 温差钳 >= 0 [K]
FC_DL_ClinkerCoolingRateCalc := xValid;                                            // 返回码：TRUE = 计算可信

END_FUNCTION

(* ---- FC_DL_CoagDoseFromJarTest.st ---- *)
(*
  道莅工业代码库 / Daoli Industrial ST Library
  组件: FC_DL_CoagDoseFromJarTest
  分类: DL_Process
  开源溯源: 无（clean-room 工程公式自研；参考公开工艺计算公式，未复制任何受版权保护代码）
  许可证: 本项目自有 (MIT)
  功能: 由烧杯试验最佳投加量反算混凝剂计量泵体积流量 [L/h]，含母液浓度换算、人工修正与上限饱和
*)
FUNCTION FC_DL_CoagDoseFromJarTest : BOOL
VAR_INPUT
    rJarDoseMgL : REAL; // 罐试最佳投加量（以进水体积计）[mg/L] / jar-test optimum dose per litre of raw water
    rFlowM3h : REAL; // 处理水量 [m3/h] / treated water flow
    rDoseTrim : REAL; // 人工修正系数 [1]，1.0 = 不修正 / manual trim factor, 1.0 = no trim
    rDoseMaxLh : REAL; // 计量泵投加体积上限 [L/h] / dosing pump volumetric upper limit
    rStockGL : REAL; // 母液有效浓度 [g/L] / stock solution effective concentration
END_VAR
VAR_OUTPUT
    rDoseLh : REAL; // 投加体积流量 [L/h] / dosing volumetric flow
    bValid : BOOL; // 结果有效位 [-] / result valid flag
    iErrCode : INT; // 事件码 0=正常 1=母液浓度非法 2=水量非法 3=超上限饱和 4=结果非有限 / event code
END_VAR
VAR
    rDoseGh : REAL; // 药剂质量流量中间量 [g/h] / intermediate coagulant mass flow
END_VAR

    // —— 段 0：全路径预清 —— //
    rDoseGh := 0.0;
    rDoseLh := 0.0;
    bValid := FALSE;
    iErrCode := 0;
    FC_DL_CoagDoseFromJarTest := FALSE;
    // —— 段 1：分母闸（母液浓度、水量） —— //
    IF ABS(rStockGL) <= 1.0E-9 THEN
        iErrCode := 1; // 母液浓度非法，无法由质量流量换算体积流量 / bad stock concentration, volume flow not derivable
        RETURN;
    END_IF;
    IF rFlowM3h <= 0.0 THEN
        iErrCode := 2; // 无处理水量，投加量保持零 / no water flow, dose held at zero
        RETURN;
    END_IF;
    // —— 段 2：量纲链 (mg/L)*(m3/h) = (g/m3)*(m3/h) = g/h；再 /(g/L) 得 L/h —— //
    rDoseGh := rJarDoseMgL * rFlowM3h; // 药剂质量流量 [g/h] / coagulant mass flow
    rDoseLh := rDoseGh / rStockGL * rDoseTrim; // 投加体积流量 [L/h] / dosing volumetric flow
    // —— 段 3：结果域闸（非有限即归零） —— //
    IF ABS(rDoseLh) > 1.0E15 THEN
        rDoseLh := 0.0;
        iErrCode := 4; // 结果非有限，强制归零 / non-finite result, forced to zero
        RETURN;
    END_IF;
    // —— 段 4：限幅 [0, rDoseMaxLh]，负值归零、超上限饱和并置码 —— //
    IF rDoseLh < 0.0 THEN
        rDoseLh := 0.0; // 负投加无物理意义 / negative dose is unphysical
    END_IF;
    IF rDoseLh > rDoseMaxLh THEN
        rDoseLh := MAX(rDoseMaxLh, 0.0); // 饱和到泵上限（上限为负时取零）/ saturate to pump limit, floor zero
        iErrCode := 3; // 信息级：超上限已饱和 / info level: saturated at upper limit
    END_IF;
    bValid := TRUE;
    FC_DL_CoagDoseFromJarTest := TRUE;
END_FUNCTION

(* ---- FC_DL_CoagulantDoseCalc.st ---- *)
(*
  ============================================================
  组件名 : FC_DL_CoagulantDoseCalc
  分类   : DL_Process
  功能   : 混凝剂投加量计算，按浊度比例前馈放大基准投加率并限幅后折算小时投加量
  开源溯源 : internal-design（本轮无外部代码逐行引用）
             参考语义 : 无外部参考
  复杂度 : C1
  版本   : 1.0.0
  ============================================================
*)

FUNCTION FC_DL_CoagulantDoseCalc : REAL
VAR_INPUT
    rFlow_m3h        : REAL; // 处理水量 [m3/h] treated water flow [m3 per hour]
    rTurbidity_Ntu   : REAL; // 实测原水浊度 [NTU] measured raw water turbidity [NTU]
    rTurbidityRef    : REAL; // 基准浊度 [NTU] reference turbidity [NTU]
    rDoseRef_mgL     : REAL; // 基准投加率 [mg/L] reference dose [mg per litre]
    rDoseMax_mgL     : REAL; // 投加率上限 [mg/L] dose ceiling [mg per litre]
    rDoseMin_mgL     : REAL; // 投加率下限 [mg/L] dose floor [mg per litre]
END_VAR
VAR_OUTPUT
    rDose_mgL     : REAL; // 实际投加率 [mg/L] applied dose [mg per litre]
    rDoseRate_kgh : REAL; // 小时投加量 [kg/h] hourly dosing rate [kg per hour]
    bValid        : BOOL; // 结果有效标志 result validity flag
END_VAR
VAR CONSTANT
    DL_MG_PER_KG : REAL := 1000.0; // 每千克毫克数 milligrams per kilogram
    DL_EPS_R     : REAL := 1.0E-6; // 实数零判定阈值 real zero threshold
END_VAR
VAR
    _bFin  : BOOL := FALSE; // 五实数输入有限性判定 finiteness verdict of the five real inputs
    _rRaw  : REAL := 0.0; // 前馈投加率 [mg/L] feed forward dose [mg per litre]
    _rDose : REAL := 0.0; // 限幅后的投加率 [mg/L] limited dose [mg per litre]
    _rLo   : REAL := 0.0; // 限幅下限 [mg/L] lower limit [mg per litre]
    _rHi   : REAL := 0.0; // 限幅上限 [mg/L] upper limit [mg per litre]
    _rRate : REAL := 0.0; // 小时投加量中间量 [kg/h] intermediate hourly rate [kg per hour]
END_VAR

// 段 1｜出口预置 preset the exit
FC_DL_CoagulantDoseCalc := 0.0; // 缺省返回零 default zero return
rDose_mgL := 0.0; // 投加率预置零 dose preset to zero
rDoseRate_kgh := 0.0; // 小时投加量预置零 hourly rate preset to zero
bValid := FALSE; // 计算完成前不认结果 unusable before the calculation
// 段 2｜非有限闸 finiteness gate
_bFin := (rFlow_m3h = rFlow_m3h) AND (rTurbidity_Ntu = rTurbidity_Ntu) AND (rTurbidityRef = rTurbidityRef) AND (rDoseRef_mgL = rDoseRef_mgL) AND (rDoseMax_mgL = rDoseMax_mgL) AND (rDoseMin_mgL = rDoseMin_mgL); // 六输入自反判定 self comparison of the six inputs
IF NOT _bFin THEN
    RETURN; // 非有限即无效 non finite means invalid
END_IF
// 段 3｜基准与流量闸 reference and flow gate
IF (rTurbidityRef <= DL_EPS_R) OR (rFlow_m3h < 0.0) OR (rTurbidity_Ntu < 0.0) OR (rDoseRef_mgL < 0.0) THEN
    RETURN; // 基准浊度非正或负流量负浊度 an illegal reference turbidity flow or dose
END_IF
// 段 4｜前馈投加率与限幅 feed forward dose and the limitation
_rRaw := rDoseRef_mgL * (rTurbidity_Ntu / rTurbidityRef); // 按浊度比例前馈 scale the dose by the turbidity ratio
_rLo := rDoseMin_mgL; // 取下限 take the floor
_rHi := rDoseMax_mgL; // 取上限 take the ceiling
IF _rLo > _rHi THEN
    _rLo := rDoseMax_mgL; // 上下限倒置时下限取原上限 an inverted pair swaps the floor
    _rHi := rDoseMin_mgL; // 上下限倒置时上限取原下限 an inverted pair swaps the ceiling
END_IF
IF _rLo < 0.0 THEN
    _rLo := 0.0; // 负下限按零处理 a negative floor becomes zero
END_IF
_rDose := LIMIT(_rLo, _rRaw, _rHi); // 限幅到上下限之间 limit the dose between the bounds
rDose_mgL := _rDose; // 投加率落定 land the dose
// 段 5｜小时投加量与出口 hourly rate and the exit
_rRate := _rDose * rFlow_m3h / DL_MG_PER_KG; // 浓度乘流量折千克 hourly mass from the dose and the flow
rDoseRate_kgh := _rRate; // 小时投加量落定 land the hourly rate
bValid := TRUE; // 结果可用 result usable
FC_DL_CoagulantDoseCalc := _rDose; // 函数返回投加率 return the dose
END_FUNCTION

(* ---- FC_DL_CoaterArealLoadingCalc.st ---- *)
(*
  Name: FC_DL_CoaterArealLoadingCalc
  Category: DL_Process
  Version: 1.0.0
  Round: R90 / 2026-11-25
  开源溯源：clean-room 自研（族 锂电极片涂布辊压，ST 开源生态实测 0 命中，无外部代码引入）
  功能：1) 由干膜厚度与涂层密度算面密度：面密度 = 厚度 × 密度，
           单位换算后为 mg/cm2。推导：厚度 µm × 密度 g/cm3 得 mg/cm2 需先除 10，
           因为 1 µm × 1 g/cm3 = 1e-4 cm × 1 g/cm3 = 1e-4 g/cm2 = 0.1 mg/cm2，
           故 fArealMgCm2 = fDryThickUm × fDensityGcm3 / 10。
        2) 与目标面密度比较给出相对偏差 fDevPct = (实测 − 目标) / 目标 × 100，
           方向为「实测减目标」：正值表示超涂（面密度偏高），负值表示欠涂。
           偏差绝对值不超过容差 fTolPct 则判合格 xPass。
  边界条件：1) 非有限值闸：四路实值入参统一过 NOT(x > -DL_BIG AND x < DL_BIG)，
           同时拦 NaN 与 Inf，命中即拦断实值通路（两个 REAL 输出强制 0.0、xPass 强制 FALSE）
           并置无效（R19），无效数据不得判合格。
        2) 分母零闸：ABS(fTargetMgCm2) > DL_EPS 才允许算相对偏差（目标为 0 时相对偏差无定义），
           否则判无效；厚度为 0 属合法工况（未涂布），面密度 0，但相对偏差仍可算。
        3) 负值闸：干膜厚度为负、密度为负、目标面密度为负、容差为负均判无效
           （容差为负会使合格判据恒假，属组态错误）。
        4) 容差窄闸：fTolPct 钳 0 ~ 100 %，越域判无效；容差为 0 表示零公差（严判），属合法组态。
        5) 饱和钳制：面密度钳 0 ~ DL_AREAL_MAX(1000 mg/cm2)，偏差钳 −1000 ~ +1000 %，
           防极端输入溢出。
  量纲自证：fArealMgCm2 = µm × (g/cm3) / 10 (mg/cm2 per µm·g/cm3) = mg/cm2，量纲闭合；
           fDevPct = (mg/cm2 − mg/cm2) / (mg/cm2) × 100 = 无因次百分数 [%]，
           分子分母同量纲，减法两侧同量纲。
*)

FUNCTION FC_DL_CoaterArealLoadingCalc : BOOL
VAR_INPUT
    fDryThickUm   : REAL;   // 干膜厚度 [µm] / Dry film thickness [µm]
    fDensityGcm3  : REAL;   // 涂层压实密度 [g/cm3] / Coating density [g/cm3]
    fTargetMgCm2  : REAL;   // 目标面密度 [mg/cm2] / Target areal loading [mg/cm2]
    fTolPct       : REAL;   // 面密度容差 [%] / Areal loading tolerance [%]
END_VAR
VAR_OUTPUT
    fArealMgCm2   : REAL;   // 实测面密度 [mg/cm2] / Measured areal loading [mg/cm2]
    fDevPct       : REAL;   // 相对偏差（实测 − 目标）[%] / Relative deviation [%]
    xPass         : BOOL;   // 面密度合格标志 [bool] / Areal loading pass flag [bool]
    xValid        : BOOL;   // 计算有效标志 [bool] / Calculation valid flag [bool]
END_VAR
VAR
    _fArealRaw    : REAL;   // 未饱和的面密度 [mg/cm2] / Raw areal loading [mg/cm2]
    _fDevRawPct   : REAL;   // 未饱和的相对偏差 [%] / Raw relative deviation [%]
    _fTolClampPct : REAL;   // 钳制后的容差 [%] / Clamped tolerance [%]
END_VAR
VAR CONSTANT
    DL_EPS        : REAL := 1.0E-9;    // 分母零闸阈值 [-] / Division-zero gate threshold [-]
    DL_BIG        : REAL := 1.0E12;    // 非有限值闸量级上限 [-] / Finiteness gate magnitude [-]
    DL_PCT        : REAL := 100.0;     // 百分比换算因子 [%] / Percent conversion factor [%]
    DL_UM_TO_MGCM2: REAL := 10.0;      // µm·g/cm3 → mg/cm2 的除数 [-] / Thickness-density divisor [-]
    DL_AREAL_MAX  : REAL := 1000.0;    // 面密度饱和上限 [mg/cm2] / Areal loading saturation ceiling
    DL_DEV_MAX    : REAL := 1000.0;    // 偏差饱和上限 [%] / Deviation saturation ceiling [%]
END_VAR

(* —— 段 1：非有限值闸（R19：四路入参全覆盖，拦 NaN 与 Inf） —— *)
IF NOT (fDryThickUm > -DL_BIG AND fDryThickUm < DL_BIG)
   OR NOT (fDensityGcm3 > -DL_BIG AND fDensityGcm3 < DL_BIG)
   OR NOT (fTargetMgCm2 > -DL_BIG AND fTargetMgCm2 < DL_BIG)
   OR NOT (fTolPct > -DL_BIG AND fTolPct < DL_BIG) THEN
    fArealMgCm2 := 0.0;                     // 输出强制 0.0 / Output forced to zero
    fDevPct := 0.0;                         // 偏差强制 0.0 / Deviation forced to zero
    xPass := FALSE;                         // 合格标志强制 FALSE / Pass forced off
    xValid := FALSE;                        // 有效位清零 / Validity cleared
    FC_DL_CoaterArealLoadingCalc := FALSE;  // 返回码同源 / Return mirrors validity
    RETURN;                                 // 立即退出 / Immediate exit
END_IF

(* —— 段 2：分母零闸（R4：目标面密度是相对偏差的分母） —— *)
IF ABS(fTargetMgCm2) <= DL_EPS THEN
    fArealMgCm2 := 0.0;                     // 输出强制 0.0 / Output forced to zero
    fDevPct := 0.0;                         // 偏差强制 0.0 / Deviation forced to zero
    xPass := FALSE;                         // 合格标志强制 FALSE / Pass forced off
    xValid := FALSE;                        // 判无效 / Invalid
    FC_DL_CoaterArealLoadingCalc := FALSE;  // 返回码同步 / Return synchronised
    RETURN;                                 // 提前退出 / Early exit
END_IF

(* —— 段 3：负值闸（负容差会使合格判据恒假，属组态错误） —— *)
IF (fDryThickUm < 0.0) OR (fDensityGcm3 < 0.0) OR (fTargetMgCm2 < 0.0) OR (fTolPct < 0.0) THEN
    fArealMgCm2 := 0.0;                     // 输出强制 0.0 / Output forced to zero
    fDevPct := 0.0;                         // 偏差强制 0.0 / Deviation forced to zero
    xPass := FALSE;                         // 合格标志强制 FALSE / Pass forced off
    xValid := FALSE;                        // 判无效 / Invalid
    FC_DL_CoaterArealLoadingCalc := FALSE;  // 返回码同步 / Return synchronised
    RETURN;                                 // 提前退出 / Early exit
END_IF

(* —— 段 4：面密度主算式（R22 方向自核：厚度乘密度，除 10 做单位换算） —— *)
_fArealRaw := fDryThickUm * fDensityGcm3 / DL_UM_TO_MGCM2;       // [mg/cm2]

(* —— 段 5：相对偏差（分子方向：实测减目标，正值 = 超涂） —— *)
_fDevRawPct := (_fArealRaw - fTargetMgCm2) / fTargetMgCm2 * DL_PCT;   // [%]

(* —— 段 6：输出单点写盘（饱和钳制后判合格，保证判据与出口同源） —— *)
fArealMgCm2 := LIMIT(0.0, _fArealRaw, DL_AREAL_MAX);             // 面密度 [mg/cm2]
fDevPct := LIMIT(-DL_DEV_MAX, _fDevRawPct, DL_DEV_MAX);          // 偏差 [%]
_fTolClampPct := LIMIT(0.0, fTolPct, DL_PCT);                    // 容差钳 0..100 [%]

(* —— 段 7：有效位与合格位单点聚合 —— *)
xValid := (fDryThickUm >= 0.0) AND (fDensityGcm3 > DL_EPS)
          AND (fTargetMgCm2 > DL_EPS) AND (fTolPct <= DL_PCT);   // 有效位聚合
xPass := xValid AND (ABS(fDevPct) <= _fTolClampPct);             // 偏差绝对值不超容差即合格
FC_DL_CoaterArealLoadingCalc := xValid;                          // 返回码：TRUE = 计算可信

END_FUNCTION

(* ---- FC_DL_CoaterDryZoneHeatCalc.st ---- *)
(*
  Name: FC_DL_CoaterDryZoneHeatCalc
  Category: DL_Process
  Version: 1.0.0
  Round: R90 / 2026-11-25
  开源溯源：clean-room 自研（族 锂电极片涂布辊压，ST 开源生态实测 0 命中，无外部代码引入）
  功能：1) 烘箱溶剂蒸发所需热量按潜热折算：Q_evap[kW] = 溶剂质量流量[kg/h] × 蒸发潜热[kJ/kg]
           / 3600[s/h]，再按热效率归一化（除以效率比例），得到实际需投入的热功率。
           效率归一化的方向是「除以效率」而不是「乘效率」：效率越低，投入必须越多，
           这是本件最容易写反的一处（写成乘会把低效烘箱算成省能）。
        2) 循环风加热所需热量按显热折算：Q_air[kW] = 风量[m3/h] × 密度[kg/m3] × 定压比热[kJ/(kg·K)]
           × 设计温升[K] / 3600，其中设计温升 DL_DT_AIR 是烘箱新风加热的设计工况常数。
           两路热量互为补充：蒸发热是工艺负荷，风加热是设备热惯性负荷，合计为烘箱热负荷。
  边界条件：1) 非有限值闸：四路实值入参统一过 NOT(x > -DL_BIG AND x < DL_BIG)，
           同时拦 NaN 与 Inf，命中即拦断实值通路（两个 REAL 输出强制 0.0）并置无效（R19）。
        2) 分母零闸：热效率比例必须 ABS > DL_EPS，否则「除以效率」发散（效率为 0 表示无热输入，
           物理上无法蒸发任何溶剂）；3600 s/h 为常量，无零风险。
        3) 效率窄闸：必须落在 DL_EFF_MIN(1 %) ~ 100 %，越域钳边界算参考值但置无效；
           超过 100 % 违反热力学第一定律，属组态错误。
        4) 负值闸：溶剂流量、潜热、风量任一为负判无效（不取绝对值掩盖反向）。
        5) 零值语义：溶剂流量为 0（未涂布）属合法工况，蒸发热为 0，不判无效；
           潜热为 0 判无效（潜热是物料属性常数，为 0 表示未组态）。
        6) 饱和钳制：两路热量均钳 0 ~ DL_Q_MAX(10000 kW)，防组态越界溢出。
  量纲自证：Q_evap = (kg/h) × (kJ/kg) / (s/h) = kJ/s = kW，除效率 [-] 后仍为 kW；
           Q_air = (m3/h) × (kg/m3) × (kJ/(kg·K)) × K / (s/h) = kJ/s = kW；
           两输出同为 kW，可相加；本件未出现 kW/kW 无因次量与温度相加的混算。
*)

FUNCTION FC_DL_CoaterDryZoneHeatCalc : BOOL
VAR_INPUT
    fSolventKgH    : REAL;   // 溶剂蒸发质量流量 [kg/h] / Solvent evaporation mass flow [kg/h]
    fLatentKJkg    : REAL;   // 溶剂蒸发潜热 [kJ/kg] / Solvent latent heat of vaporization [kJ/kg]
    fEfficiencyPct : REAL;   // 烘箱热效率 [%] / Oven thermal efficiency [%]
    fAirFlowM3h    : REAL;   // 循环/新风体积流量 [m3/h] / Air volumetric flow [m3/h]
END_VAR
VAR_OUTPUT
    fHeatKW        : REAL;   // 溶剂蒸发所需热功率（已效率归一）[kW] / Evaporation heat demand [kW]
    fAirHeatKW     : REAL;   // 风加热所需热功率 [kW] / Air heating heat demand [kW]
    fTotalKW       : REAL;   // 烘箱总热负荷 [kW] / Total oven heat load [kW]
    xValid         : BOOL;   // 计算有效标志 [bool] / Calculation valid flag [bool]
END_VAR
VAR
    _fEffRatio     : REAL;   // 归一化热效率 [-] / Normalized thermal efficiency [-]
    _fEvapRawKW    : REAL;   // 未效率归一的蒸发热功率 [kW] / Raw evaporation heat [kW]
    _fHeatRawKW    : REAL;   // 效率归一后的蒸发热功率 [kW] / Efficiency-normalized heat [kW]
    _fAirRawKW     : REAL;   // 未饱和的风加热功率 [kW] / Raw air heating heat [kW]
END_VAR
VAR CONSTANT
    DL_EPS         : REAL := 1.0E-9;    // 分母零闸阈值 [-] / Division-zero gate threshold [-]
    DL_BIG         : REAL := 1.0E12;    // 非有限值闸量级上限 [-] / Finiteness gate magnitude [-]
    DL_PCT         : REAL := 100.0;     // 百分比换算因子 [%] / Percent conversion factor [%]
    DL_S_PER_H     : REAL := 3600.0;    // h → s 换算因子 [s/h] / Hour to second factor [s/h]
    DL_RHO_AIR     : REAL := 1.20;      // 空气密度 [kg/m3] / Air density [kg/m3]
    DL_CP_AIR      : REAL := 1.005;     // 空气定压比热 [kJ/(kg·K)] / Air specific heat [kJ/(kg·K)]
    DL_DT_AIR      : REAL := 100.0;     // 烘箱设计温升 [K] / Oven design temperature rise [K]
    DL_EFF_MIN     : REAL := 1.0;       // 热效率下限 [%] / Thermal efficiency lower bound [%]
    DL_Q_MAX       : REAL := 10000.0;   // 热功率饱和上限 [kW] / Heat power saturation ceiling [kW]
END_VAR

(* —— 段 1：非有限值闸（R19：四路入参全覆盖，拦 NaN 与 Inf） —— *)
IF NOT (fSolventKgH > -DL_BIG AND fSolventKgH < DL_BIG)
   OR NOT (fLatentKJkg > -DL_BIG AND fLatentKJkg < DL_BIG)
   OR NOT (fEfficiencyPct > -DL_BIG AND fEfficiencyPct < DL_BIG)
   OR NOT (fAirFlowM3h > -DL_BIG AND fAirFlowM3h < DL_BIG) THEN
    fHeatKW := 0.0;                         // 输出强制 0.0 / Output forced to zero
    fAirHeatKW := 0.0;                      // 风加热强制 0.0 / Air heat forced to zero
    fTotalKW := 0.0;                        // 总负荷强制 0.0 / Total load forced to zero
    xValid := FALSE;                        // 有效位清零 / Validity cleared
    FC_DL_CoaterDryZoneHeatCalc := FALSE;   // 返回码同源 / Return mirrors validity
    RETURN;                                 // 立即退出 / Immediate exit
END_IF

(* —— 段 2：分母零闸（R4：热效率是除数，为 0 则需热量发散） —— *)
IF ABS(fEfficiencyPct / DL_PCT) <= DL_EPS THEN
    fHeatKW := 0.0;                         // 输出强制 0.0 / Output forced to zero
    fAirHeatKW := 0.0;                      // 风加热强制 0.0 / Air heat forced to zero
    fTotalKW := 0.0;                        // 总负荷强制 0.0 / Total load forced to zero
    xValid := FALSE;                        // 判无效 / Invalid
    FC_DL_CoaterDryZoneHeatCalc := FALSE;   // 返回码同步 / Return synchronised
    RETURN;                                 // 提前退出 / Early exit
END_IF

(* —— 段 3：负值闸（流量与潜热均不可为负） —— *)
IF (fSolventKgH < 0.0) OR (fLatentKJkg < 0.0) OR (fAirFlowM3h < 0.0) THEN
    fHeatKW := 0.0;                         // 输出强制 0.0 / Output forced to zero
    fAirHeatKW := 0.0;                      // 风加热强制 0.0 / Air heat forced to zero
    fTotalKW := 0.0;                        // 总负荷强制 0.0 / Total load forced to zero
    xValid := FALSE;                        // 判无效 / Invalid
    FC_DL_CoaterDryZoneHeatCalc := FALSE;   // 返回码同步 / Return synchronised
    RETURN;                                 // 提前退出 / Early exit
END_IF

(* —— 段 4：蒸发热功率（R22 方向自核：效率在分母，效率越低投入越大） —— *)
_fEvapRawKW := fSolventKgH * fLatentKJkg / DL_S_PER_H;            // 理论蒸发热 [kW]
_fEffRatio := LIMIT(DL_EFF_MIN, fEfficiencyPct, DL_PCT) / DL_PCT; // 效率归一，并钳到 1~100 %
_fHeatRawKW := _fEvapRawKW / _fEffRatio;                          // 效率归一后热功率 [kW]

(* —— 段 5：风加热功率（显热式：风量 × 密度 × 比热 × 温升，除 3600 得 kW） —— *)
_fAirRawKW := fAirFlowM3h * DL_RHO_AIR * DL_CP_AIR * DL_DT_AIR / DL_S_PER_H;   // [kW]

(* —— 段 6：输出单点写盘（饱和钳制后合计，保证合计值取自同一组出口值） —— *)
fHeatKW := LIMIT(0.0, _fHeatRawKW, DL_Q_MAX);                     // 蒸发热需求 [kW]
fAirHeatKW := LIMIT(0.0, _fAirRawKW, DL_Q_MAX);                   // 风加热需求 [kW]
fTotalKW := LIMIT(0.0, fHeatKW + fAirHeatKW, DL_Q_MAX);           // 总热负荷 [kW]

(* —— 段 7：有效位单点聚合（效率窄闸 + 潜热已组态 + 风量非负） —— *)
xValid := (fEfficiencyPct >= DL_EFF_MIN) AND (fEfficiencyPct <= DL_PCT)   // 效率在 1..100 %
          AND (fLatentKJkg > DL_EPS)                                      // 潜热已组态
          AND (fSolventKgH >= 0.0)                                        // 溶剂流量非负
          AND (fAirFlowM3h >= 0.0);                                       // 风量非负
FC_DL_CoaterDryZoneHeatCalc := xValid;                            // 返回码：TRUE = 计算可信

END_FUNCTION

(* ---- FC_DL_CoaterSolventBalanceCalc.st ---- *)
(*
  Name: FC_DL_CoaterSolventBalanceCalc
  Category: DL_Process
  Version: 1.0.0
  Round: R90 / 2026-11-25
  开源溯源：clean-room 自研（族 锂电极片涂布辊压，ST 开源生态实测 0 命中，无外部代码引入）
  功能：1) 溶剂衡算按「入料带入 − 烘干排出 = 残留」建立：湿涂层质量流量乘以浆料溶剂比例得到
           入料带入的溶剂量，减去排风侧实测带走的溶剂量，差值即留在极片中的残留溶剂量。
           差值的符号口径固定为「带入减排出」：正值 = 有残留（正常），负值 = 排出大于带入
           （物料不平衡，通常是排风侧传感器偏高或入料计量偏低）。
        2) 残留比例 = 残留量 / 带入量 × 100，与残留上限 fResidualLimitPct 比较给出超限标志 xOver。
           比例的分母是「带入量」而不是「排出量」或「湿涂层总量」：判据语义是
           「有多少比例的溶剂没被烘干」，故必须以带入量为基准。
  边界条件：1) 非有限值闸：四路实值入参统一过 NOT(x > -DL_BIG AND x < DL_BIG)，
           同时拦 NaN 与 Inf，命中即拦断实值通路（两个 REAL 输出强制 0.0、xOver 强制 FALSE）
           并置无效（R19），无效数据不得判超限。
        2) 分母零闸：带入溶剂量（fCoatingKgH × fSolventPct/100）必须 ABS > DL_EPS，
           否则残留比例无定义；带入量为 0 表示未涂布，判无效而不输出比例。
        3) 溶剂比例窄闸：fSolventPct 必须落在 0 ~ 100 %，越域钳边界并置无效（超过 100 % 不可能）。
        4) 物料不平衡闸：排出量大于带入量时，差值物理上不可能为正残留，故残留量钳 0、
           残留比例钳 0，并置 xValid=FALSE 上报物料不平衡（不输出负残留掩盖问题）。
        5) 负值闸：涂层质量流量、排出量、上限比例任一为负判无效。
        6) 饱和钳制：残留量钳 0 ~ DL_RES_MAX(10000 kg/h)，残留比例钳 0 ~ 100 %。
  量纲自证：入料带入 = (kg/h) × (%/100) = kg/h；残留 = (kg/h) − (kg/h) = kg/h，减法同量纲；
           残留比例 = (kg/h) / (kg/h) × 100 = 无因次百分数 [%]，与上限比例同量纲；
           本件未出现 kg/h 与 % 直接相加的混算。
*)

FUNCTION FC_DL_CoaterSolventBalanceCalc : BOOL
VAR_INPUT
    fCoatingKgH      : REAL;   // 湿涂层质量流量 [kg/h] / Wet coating mass flow [kg/h]
    fSolventPct      : REAL;   // 浆料溶剂质量比例 [%] / Slurry solvent mass ratio [%]
    fExhaustKgH      : REAL;   // 排风带走溶剂量 [kg/h] / Solvent removed by exhaust [kg/h]
    fResidualLimitPct: REAL;   // 残留溶剂上限 [%] / Residual solvent upper limit [%]
END_VAR
VAR_OUTPUT
    fResidualKgH     : REAL;   // 残留溶剂量 [kg/h] / Residual solvent mass flow [kg/h]
    fResidualPct     : REAL;   // 残留溶剂比例 [%] / Residual solvent ratio [%]
    xOver            : BOOL;   // 残留超限标志 [bool] / Residual over-limit flag [bool]
    xValid           : BOOL;   // 计算有效标志 [bool] / Calculation valid flag [bool]
END_VAR
VAR
    _fSolventRatio   : REAL;   // 归一化溶剂比例 [-] / Normalized solvent ratio [-]
    _fSolventInKgH   : REAL;   // 入料带入溶剂量 [kg/h] / Solvent carried in by coating [kg/h]
    _fResidualRaw    : REAL;   // 未钳制的残留量（可能为负）[kg/h] / Raw residual, may be negative [kg/h]
    _fResidualClamp  : REAL;   // 钳制后的残留量 [kg/h] / Clamped residual [kg/h]
    _fPctRaw         : REAL;   // 未饱和的残留比例 [%] / Raw residual ratio [%]
    _bBalanceOk      : BOOL;   // 物料平衡合法（排出不超过带入）[bool] / Mass balance valid [bool]
END_VAR
VAR CONSTANT
    DL_EPS           : REAL := 1.0E-9;    // 分母零闸阈值 [-] / Division-zero gate threshold [-]
    DL_BIG           : REAL := 1.0E12;    // 非有限值闸量级上限 [-] / Finiteness gate magnitude [-]
    DL_PCT           : REAL := 100.0;     // 百分比换算因子 [%] / Percent conversion factor [%]
    DL_RES_MAX       : REAL := 10000.0;   // 残留量饱和上限 [kg/h] / Residual saturation ceiling [kg/h]
END_VAR

(* —— 段 1：非有限值闸（R19：四路入参全覆盖，拦 NaN 与 Inf） —— *)
IF NOT (fCoatingKgH > -DL_BIG AND fCoatingKgH < DL_BIG)
   OR NOT (fSolventPct > -DL_BIG AND fSolventPct < DL_BIG)
   OR NOT (fExhaustKgH > -DL_BIG AND fExhaustKgH < DL_BIG)
   OR NOT (fResidualLimitPct > -DL_BIG AND fResidualLimitPct < DL_BIG) THEN
    fResidualKgH := 0.0;                    // 输出强制 0.0 / Output forced to zero
    fResidualPct := 0.0;                    // 比例强制 0.0 / Ratio forced to zero
    xOver := FALSE;                         // 超限强制 FALSE / Over-limit forced off
    xValid := FALSE;                        // 有效位清零 / Validity cleared
    FC_DL_CoaterSolventBalanceCalc := FALSE;   // 返回码同源 / Return mirrors validity
    RETURN;                                 // 立即退出 / Immediate exit
END_IF

(* —— 段 2：负值闸（流量与上限比例均不可为负） —— *)
IF (fCoatingKgH < 0.0) OR (fExhaustKgH < 0.0) OR (fResidualLimitPct < 0.0) THEN
    fResidualKgH := 0.0;                    // 输出强制 0.0 / Output forced to zero
    fResidualPct := 0.0;                    // 比例强制 0.0 / Ratio forced to zero
    xOver := FALSE;                         // 超限强制 FALSE / Over-limit forced off
    xValid := FALSE;                        // 判无效 / Invalid
    FC_DL_CoaterSolventBalanceCalc := FALSE;   // 返回码同步 / Return synchronised
    RETURN;                                 // 提前退出 / Early exit
END_IF

(* —— 段 3：带入溶剂量与分母零闸（R4：带入量是残留比例的分母） —— *)
_fSolventRatio := LIMIT(0.0, fSolventPct, DL_PCT) / DL_PCT;       // 溶剂比例归一并钳 0..100 %
_fSolventInKgH := fCoatingKgH * _fSolventRatio;                   // 入料带入溶剂量 [kg/h]
IF ABS(_fSolventInKgH) <= DL_EPS THEN
    fResidualKgH := 0.0;                    // 输出强制 0.0 / Output forced to zero
    fResidualPct := 0.0;                    // 比例强制 0.0 / Ratio forced to zero
    xOver := FALSE;                         // 超限强制 FALSE / Over-limit forced off
    xValid := FALSE;                        // 判无效 / Invalid
    FC_DL_CoaterSolventBalanceCalc := FALSE;   // 返回码同步 / Return synchronised
    RETURN;                                 // 提前退出 / Early exit
END_IF

(* —— 段 4：衡算主算式（R22 符号方向自核：带入减排出，正值 = 有残留） —— *)
_fResidualRaw := _fSolventInKgH - fExhaustKgH;                    // 残留量 [kg/h]（可能为负）
_bBalanceOk := (_fResidualRaw >= 0.0);                            // 物料平衡合法性
_fResidualClamp := MAX(0.0, _fResidualRaw);                       // 负残留钳 0，不输出负值
_fPctRaw := _fResidualClamp / _fSolventInKgH * DL_PCT;            // 残留比例 [%]

(* —— 段 5：输出单点写盘（饱和钳制后判超限，保证判据与出口同源） —— *)
fResidualKgH := LIMIT(0.0, _fResidualClamp, DL_RES_MAX);          // 残留量 [kg/h]
fResidualPct := LIMIT(0.0, _fPctRaw, DL_PCT);                     // 残留比例钳 0..100 [%]

(* —— 段 6：有效位单点聚合（溶剂比例窄闸 + 物料平衡 + 带入量可归一） —— *)
xValid := (fSolventPct >= 0.0) AND (fSolventPct <= DL_PCT)        // 溶剂比例在 0..100 %
          AND (_bBalanceOk)                                       // 排出不得超过带入
          AND (_fSolventInKgH > DL_EPS);                          // 带入量可作分母

(* —— 段 7：超限判定（无效数据不得判超限） —— *)
xOver := xValid AND (fResidualPct > fResidualLimitPct);
FC_DL_CoaterSolventBalanceCalc := xValid;                         // 返回码：TRUE = 计算可信

END_FUNCTION

(* ---- FC_DL_CoaterTensionZoneCalc.st ---- *)
(*
  Name: FC_DL_CoaterTensionZoneCalc
  Category: DL_Process
  Version: 1.0.0
  Round: R90 / 2026-11-25
  开源溯源：clean-room 自研（族 锂电极片涂布辊压，ST 开源生态实测 0 命中，无外部代码引入）
  功能：1) 分区总张力按「幅宽 × 单位宽度张力」计算：fTensionN = 幅宽[mm] × 单位张力[N/mm]。
           单位宽度张力是涂布机张力控制的标准口语口径（N/mm），乘幅宽即得该区的总张力设定值，
           幅宽变化时必须同步换算，不能沿用固定总张力（否则单位张力随幅宽漂移）。
        2) 辊面线压按「总张力摊到包角对应的接触弧长」计算：
             接触弧长 = 包角 × 辊半径 = DL_WRAP_RAD × (辊径/2)   [mm]
             辊面线压 = 总张力[N] / 接触弧长[mm]                  [N/mm]
           该口径的含义是「辊面单位母线长度承受的平均法向线压」，用于辊子刚度与轴承选型校核。
           归一化口径在此声明：分母是接触弧长（含辊径），不是幅宽、不是辊径本身，
           若改用幅宽会得到一个与单位张力完全相同的量（信息量为零），这是必须避免的写法。
  边界条件：1) 非有限值闸：三路实值入参统一过 NOT(x > -DL_BIG AND x < DL_BIG)，
           同时拦 NaN 与 Inf，命中即拦断实值通路（两个 REAL 输出强制 0.0）并置无效（R19）。
        2) 分母零闸：幅宽必须 ABS > DL_EPS（总张力按幅宽换算，幅宽为 0 无意义）；
           辊径经 DL_DIA_MIN_MM(1 mm) 下限钳制后参与接触弧长计算，防辊径为 0 使弧长为 0 而除零。
        3) 负值闸：幅宽、单位张力、辊径任一为负判无效（不取绝对值掩盖反向）。
        4) 饱和钳制：总张力钳 0 ~ DL_TEN_MAX(100000 N)、线压钳 0 ~ DL_PRESS_MAX(1000 N/mm)，
           防极端幅宽与辊径组合溢出。
  量纲自证：fTensionN = mm × (N/mm) = N；
           接触弧长 = [-] × mm = mm（包角为无因次弧度）；
           fLinePressNmm = N / mm = N/mm，与总张力量纲不同且各自自洽，未混算。
*)

FUNCTION FC_DL_CoaterTensionZoneCalc : BOOL
VAR_INPUT
    fWebWidthMm    : REAL;   // 极片幅宽 [mm] / Web width [mm]
    fUnitTensionNmm: REAL;   // 单位宽度张力 [N/mm] / Tension per unit width [N/mm]
    fRollDiaMm     : REAL;   // 导辊直径 [mm] / Roller diameter [mm]
END_VAR
VAR_OUTPUT
    fTensionN      : REAL;   // 分区总张力 [N] / Zone total tension [N]
    fLinePressNmm  : REAL;   // 辊面平均线压 [N/mm] / Mean roller face line pressure [N/mm]
    xValid         : BOOL;   // 计算有效标志 [bool] / Calculation valid flag [bool]
END_VAR
VAR
    _fTensionRawN  : REAL;   // 未饱和的总张力 [N] / Raw total tension [N]
    _fDiaClampMm   : REAL;   // 钳制后的辊径 [mm] / Clamped roller diameter [mm]
    _fArcLenMm     : REAL;   // 包角对应的接触弧长 [mm] / Contact arc length [mm]
    _fPressRawNmm  : REAL;   // 未饱和的辊面线压 [N/mm] / Raw roller line pressure [N/mm]
END_VAR
VAR CONSTANT
    DL_EPS         : REAL := 1.0E-9;    // 分母零闸阈值 [-] / Division-zero gate threshold [-]
    DL_BIG         : REAL := 1.0E12;    // 非有限值闸量级上限 [-] / Finiteness gate magnitude [-]
    DL_PI          : REAL := 3.14159265;   // 圆周率 [-] / Pi [-]
    DL_DIA_MIN_MM  : REAL := 1.0;       // 辊径下限钳制值 [mm] / Roller diameter lower clamp [mm]
    DL_TWO         : REAL := 2.0;       // 半径除数 [-] / Radius divisor [-]
    DL_TEN_MAX     : REAL := 100000.0;  // 总张力饱和上限 [N] / Total tension saturation ceiling [N]
    DL_PRESS_MAX   : REAL := 1000.0;    // 辊面线压饱和上限 [N/mm] / Line pressure saturation ceiling [N/mm]
END_VAR

(* —— 段 1：非有限值闸（R19：三路入参全覆盖，拦 NaN 与 Inf） —— *)
IF NOT (fWebWidthMm > -DL_BIG AND fWebWidthMm < DL_BIG)
   OR NOT (fUnitTensionNmm > -DL_BIG AND fUnitTensionNmm < DL_BIG)
   OR NOT (fRollDiaMm > -DL_BIG AND fRollDiaMm < DL_BIG) THEN
    fTensionN := 0.0;                       // 输出强制 0.0 / Output forced to zero
    fLinePressNmm := 0.0;                   // 线压强制 0.0 / Line pressure forced to zero
    xValid := FALSE;                        // 有效位清零 / Validity cleared
    FC_DL_CoaterTensionZoneCalc := FALSE;   // 返回码同源 / Return mirrors validity
    RETURN;                                 // 立即退出 / Immediate exit
END_IF

(* —— 段 2：分母零闸（R4：幅宽是总张力的换算基准） —— *)
IF ABS(fWebWidthMm) <= DL_EPS THEN
    fTensionN := 0.0;                       // 输出强制 0.0 / Output forced to zero
    fLinePressNmm := 0.0;                   // 线压强制 0.0 / Line pressure forced to zero
    xValid := FALSE;                        // 判无效 / Invalid
    FC_DL_CoaterTensionZoneCalc := FALSE;   // 返回码同步 / Return synchronised
    RETURN;                                 // 提前退出 / Early exit
END_IF

(* —— 段 3：负值闸（幅宽/单位张力/辊径均不可为负） —— *)
IF (fWebWidthMm < 0.0) OR (fUnitTensionNmm < 0.0) OR (fRollDiaMm < 0.0) THEN
    fTensionN := 0.0;                       // 输出强制 0.0 / Output forced to zero
    fLinePressNmm := 0.0;                   // 线压强制 0.0 / Line pressure forced to zero
    xValid := FALSE;                        // 判无效 / Invalid
    FC_DL_CoaterTensionZoneCalc := FALSE;   // 返回码同步 / Return synchronised
    RETURN;                                 // 提前退出 / Early exit
END_IF

(* —— 段 4：总张力（R22 方向自核：幅宽乘单位张力，不是除） —— *)
_fTensionRawN := fWebWidthMm * fUnitTensionNmm;                  // 总张力 [N]

(* —— 段 5：辊面线压（分母为包角接触弧长，含辊径；R22 归一化口径已在此声明） —— *)
_fDiaClampMm := MAX(DL_DIA_MIN_MM, fRollDiaMm);                  // 辊径下限钳 [mm]
_fArcLenMm := DL_PI * _fDiaClampMm / DL_TWO;                     // 180° 包角接触弧长 [mm]
_fPressRawNmm := _fTensionRawN / _fArcLenMm;                     // 辊面线压 [N/mm]

(* —— 段 6：输出单点写盘（饱和钳制） —— *)
fTensionN := LIMIT(0.0, _fTensionRawN, DL_TEN_MAX);              // 总张力 [N]
fLinePressNmm := LIMIT(0.0, _fPressRawNmm, DL_PRESS_MAX);        // 辊面线压 [N/mm]

(* —— 段 7：有效位单点聚合 —— *)
xValid := (fWebWidthMm > DL_EPS)                                 // 幅宽为正
          AND (fUnitTensionNmm >= 0.0)                          // 单位张力非负
          AND (fRollDiaMm > DL_EPS);                            // 辊径为正（弧长可算）
FC_DL_CoaterTensionZoneCalc := xValid;                           // 返回码：TRUE = 计算可信

END_FUNCTION

(* ---- FC_DL_CoaterWetThicknessCalc.st ---- *)
(*
  Name: FC_DL_CoaterWetThicknessCalc
  Category: DL_Process
  Version: 1.0.0
  Round: R90 / 2026-11-25
  开源溯源：clean-room 自研（族 锂电极片涂布辊压，ST 开源生态实测 0 命中，无外部代码引入）
  功能：1) 由目标干膜面密度与浆料固含量反算湿膜厚度，供涂布模头间隙（湿膜）设定使用。
           推导链：干燥后保留的固体质量面密度即目标面密度；湿膜中固体占质量比例为固含量，
           故湿膜质量面密度 = 干面密度 / 固含量；再由湿膜密度换算为体积厚度。
           逐步为：mg/cm2 → g/m2 乘 10；除以固含量比例得湿膜 g/m2；
           除以密度 g/cm3 直接得 µm（因为 1 g/m2 ÷ 1 g/cm3 = 1 µm，量纲恰好对消）。
        2) 固含量按百分比入参，先归一化到 0~1 再作分母，禁止直接用百分数当比例。
  边界条件：1) 非有限值闸：三路实值入参统一过 NOT(x > -DL_BIG AND x < DL_BIG)，
           同时拦 NaN 与 Inf，命中即拦断实值通路（fWetUm 强制 0.0）并置无效（R19）。
        2) 分母零闸：固含量比例必须 ABS > DL_EPS（固含量为 0 表示全溶剂，湿膜厚度趋于无穷，
           物理上不可能）；密度必须 ABS > DL_EPS（密度为 0 无意义）。
        3) 固含量窄闸：必须落在 DL_SOLID_MIN(0.1 %) ~ 100 %，越域判无效；
           上限 100 % 是「无溶剂」极限，此时湿膜 = 干膜，属合法边界值。
        4) 负值闸：面密度为负、密度为负判无效（不取绝对值掩盖反向）。
        5) 饱和钳制：湿膜厚度钳 0 ~ DL_WET_MAX(5000 µm)，防极小固含量把厚度放大到溢出。
  量纲自证：fArealMgCm2 [mg/cm2] × 10 (g/m2 per mg/cm2) = g/m2；
           除以固含量 [-]= g/m2（湿膜）；
           除以密度 [g/cm3]：g/m2 ÷ g/cm3 = cm3/m2 = 1e-6 m3/m2 = 1e-6 m = 1 µm，故结果 [µm]。
*)

FUNCTION FC_DL_CoaterWetThicknessCalc : BOOL
VAR_INPUT
    fArealMgCm2   : REAL;   // 目标干膜面密度 [mg/cm2] / Target dry areal loading [mg/cm2]
    fSolidPct     : REAL;   // 浆料固含量 [%] / Slurry solid content [%]
    fDensityGcm3  : REAL;   // 湿膜密度 [g/cm3] / Wet film density [g/cm3]
END_VAR
VAR_OUTPUT
    fWetUm        : REAL;   // 湿膜厚度 [µm] / Wet film thickness [µm]
    xValid        : BOOL;   // 计算有效标志 [bool] / Calculation valid flag [bool]
END_VAR
VAR
    _fSolidRatio  : REAL;   // 归一化固含量 [-] / Normalized solid ratio [-]
    _fDryGm2      : REAL;   // 干膜面密度 [g/m2] / Dry areal loading [g/m2]
    _fWetGm2      : REAL;   // 湿膜面密度 [g/m2] / Wet areal loading [g/m2]
    _fWetRawUm    : REAL;   // 未饱和的湿膜厚度 [µm] / Raw wet thickness [µm]
END_VAR
VAR CONSTANT
    DL_EPS        : REAL := 1.0E-9;    // 分母零闸阈值 [-] / Division-zero gate threshold [-]
    DL_BIG        : REAL := 1.0E12;    // 非有限值闸量级上限 [-] / Finiteness gate magnitude [-]
    DL_PCT        : REAL := 100.0;     // 百分比换算因子 [%] / Percent conversion factor [%]
    DL_MGCM2_TO_GM2 : REAL := 10.0;    // mg/cm2 → g/m2 换算因子 [g/m2 per mg/cm2] / Areal unit factor
    DL_SOLID_MIN  : REAL := 0.10;      // 固含量下限 [%] / Solid content lower bound [%]
    DL_WET_MAX    : REAL := 5000.0;    // 湿膜厚度饱和上限 [µm] / Wet thickness saturation ceiling [µm]
END_VAR

(* —— 段 1：非有限值闸（R19：闸断实值通路，NaN 不得进入除法链） —— *)
IF NOT (fArealMgCm2 > -DL_BIG AND fArealMgCm2 < DL_BIG)
   OR NOT (fSolidPct > -DL_BIG AND fSolidPct < DL_BIG)
   OR NOT (fDensityGcm3 > -DL_BIG AND fDensityGcm3 < DL_BIG) THEN
    fWetUm := 0.0;                          // 输出强制 0.0 / Output forced to zero
    xValid := FALSE;                        // 有效位清零 / Validity cleared
    FC_DL_CoaterWetThicknessCalc := FALSE;  // 返回码同源 / Return mirrors validity
    RETURN;                                 // 立即退出 / Immediate exit
END_IF

(* —— 段 2：分母零闸（R4：固含量与密度两个分母都必须先过 ABS 闸） —— *)
IF (ABS(fSolidPct / DL_PCT) <= DL_EPS) OR (ABS(fDensityGcm3) <= DL_EPS) THEN
    fWetUm := 0.0;                          // 输出强制 0.0 / Output forced to zero
    xValid := FALSE;                        // 判无效 / Invalid
    FC_DL_CoaterWetThicknessCalc := FALSE;  // 返回码同步 / Return synchronised
    RETURN;                                 // 提前退出 / Early exit
END_IF

(* —— 段 3：负值闸（面密度/密度为负属变送器故障，不取 ABS 掩盖） —— *)
IF (fArealMgCm2 < 0.0) OR (fDensityGcm3 < 0.0) THEN
    fWetUm := 0.0;                          // 输出强制 0.0 / Output forced to zero
    xValid := FALSE;                        // 判无效 / Invalid
    FC_DL_CoaterWetThicknessCalc := FALSE;  // 返回码同步 / Return synchronised
    RETURN;                                 // 提前退出 / Early exit
END_IF

(* —— 段 4：主算式（R22 方向自核：固含量在分母，固含量越高湿膜越薄） —— *)
_fSolidRatio := fSolidPct / DL_PCT;                              // 固含量归一 [-]
_fDryGm2 := fArealMgCm2 * DL_MGCM2_TO_GM2;                       // 干膜面密度 [g/m2]
_fWetGm2 := _fDryGm2 / _fSolidRatio;                             // 湿膜面密度 [g/m2]
_fWetRawUm := _fWetGm2 / fDensityGcm3;                           // 湿膜厚度 [µm]

(* —— 段 5：输出单点写盘（饱和钳制） —— *)
fWetUm := LIMIT(0.0, _fWetRawUm, DL_WET_MAX);                    // 湿膜厚度 [µm]

(* —— 段 6：有效位单点聚合（固含量窄闸 + 非负） —— *)
xValid := (fSolidPct >= DL_SOLID_MIN) AND (fSolidPct <= DL_PCT)  // 固含量在窄闸内
          AND (fArealMgCm2 >= 0.0)                               // 面密度非负
          AND (fDensityGcm3 > DL_EPS);                           // 密度为正
FC_DL_CoaterWetThicknessCalc := xValid;                          // 返回码：TRUE = 计算可信

END_FUNCTION

(* ---- FC_DL_CoatingPanSprayCalc.st ---- *)
(*
  DL Factory R84 | FC_DL_CoatingPanSprayCalc
  功能：按片床重量与目标增重算包衣液总量、喷射时长与回算干增重
  开源溯源：无（clean-room 自研，依据公开工艺公式，来源=行业通用公式，许可证=MIT，借鉴点=公式结构）
  规则：R1-R16 全遵守
*)
FUNCTION FC_DL_CoatingPanSprayCalc : REAL
VAR_INPUT
    fBedKg : REAL := 200.0; // 片床重量 [kg] / tablet bed mass [kg]
    fGainPct : REAL := 3.0; // 目标增重（干基） [%] / target weight gain [%]
    fSolidPct : REAL := 12.0; // 包衣液固含量 [%] / coating suspension solids [%]
    fSprayRateGmin : REAL := 120.0; // 喷量速率 [g/min] / spray rate [g/min]
    fDensityGml : REAL := 1.05; // 包衣液密度 [g/mL] / suspension density [g/mL]
END_VAR
VAR_OUTPUT
    fTotalSolL : REAL; // 包衣液总量 [L] / total suspension volume [L]
    fSprayMin : REAL; // 喷射时长 [min] / spray duration [min]
    fDryGainPct : REAL; // 回算干增重（校验用） [%] / back calculated dry gain [%]
    xValid : BOOL; // 计算结果有效标志 [-] / calculation valid flag [-]
END_VAR
VAR
    fBedG : REAL; // 片床重量折算 [g] / bed mass in grams [g]
    fDryGainG : REAL; // 目标干增重质量 [g] / target dry gain mass [g]
    fLiquidG : REAL; // 包衣液总质量（湿） [g] / total liquid mass [g]
END_VAR

// 段 1｜出口预置（R256）
FC_DL_CoatingPanSprayCalc := -1.0; // 哨兵返回 -1（无效） [-] / sentinel return -1, invalid [-]
fTotalSolL := 0.0; // 液量预置零 [L] / volume preset zero [L]
fSprayMin := 0.0; // 时长预置零 [min] / duration preset zero [min]
fDryGainPct := 0.0; // 干增重预置零 [%] / dry gain preset zero [%]
xValid := FALSE; // 计算完成前不认结果 [-] / unusable before calculation [-]

// 段 2｜非有限拦截 + 域闸（R4/R20）
IF NOT (fBedKg > -1.0E30 AND fBedKg < 1.0E30) OR NOT (fGainPct > -1.0E30 AND fGainPct < 1.0E30) OR NOT (fSolidPct > -1.0E30 AND fSolidPct < 1.0E30) OR NOT (fSprayRateGmin > -1.0E30 AND fSprayRateGmin < 1.0E30) OR NOT (fDensityGml > -1.0E30 AND fDensityGml < 1.0E30) THEN
    RETURN; // 任一入参为 NaN/Inf 一律拒绝 [-] / any NaN or Inf input rejected [-]
END_IF
IF fBedKg < 1.0E-9 OR fGainPct < 1.0E-9 OR fSolidPct < 1.0E-9 OR fSolidPct > 100.0 THEN
    RETURN; // 片床/增重/固含域闸（固含须在 (0,100]） [%] / bed, gain and solids domain gate [%]
END_IF
IF fSprayRateGmin < 1.0E-9 OR fDensityGml < 1.0E-9 THEN
    RETURN; // 喷量与密度正域分母闸（防除零） [g/min, g/mL] / spray rate and density denominator gate [-]
END_IF

// 段 3｜干增重 → 湿液量
fBedG := fBedKg * 1000.0; // kg × 1000 g/kg = g / [kg] × [g/kg] = [g]
fDryGainG := (fBedG * fGainPct) / 100.0; // g × % ÷ 100 = g / [g] × [%] / 100 = [g]
fLiquidG := (fDryGainG * 100.0) / fSolidPct; // g × 100 ÷ % = g（固含折算湿液） / [g] × 100 / [%] = [g]

// 段 4｜液量体积与喷射时长
fTotalSolL := fLiquidG / fDensityGml / 1000.0; // g ÷ g/mL = mL；mL ÷ 1000 = L / [g] / [g/mL] = [mL], [mL] / 1000 = [L]
fSprayMin := fLiquidG / fSprayRateGmin; // g ÷ g/min = min / [g] / [g/min] = [min]
IF NOT (fTotalSolL > -1.0E30 AND fTotalSolL < 1.0E30) OR NOT (fSprayMin > -1.0E30 AND fSprayMin < 1.0E30) THEN
    RETURN; // 结果非有限再拦一次 [-] / second finiteness gate on the results [-]
END_IF

// 段 5｜回算干增重（校验链：g × % ÷ g × 100 = %）
fDryGainPct := ((fLiquidG * fSolidPct) / 100.0 / fBedG) * 100.0; // [g] × [%] / [g] × 100 = [%]
xValid := TRUE; // 链路有效 [-] / chain valid [-]
FC_DL_CoatingPanSprayCalc := fSprayRateGmin; // 返回采用的喷量速率 [g/min] / return the adopted spray rate [g/min]
END_FUNCTION

(* ---- FC_DL_CompactionPressureCalc.st ---- *)
(*
  Component : FC_DL_CompactionPressureCalc
  Category  : DL_Process
  Type      : FC
  Complexity: C2
  VERSION   : v1.0.0
  功能      : 压制压力核算：按压坯相对密度与材料常数算单位压制压力，并折算压机吨位需求（含安全系数）。
  开源溯源  : 道莅原创 clean-room 自研（无外部代码引用）｜License: MIT
  边界条件  : ① 松装密度、材料常数、压制面积、安全系数须 > 1e-9，否则返回哨兵 -1；
              ② 相对密度 <= 1（压坯未致密化）时压制压力按 0 输出并置 xValid 真（合法空工况）；
              ③ 吨位折算：MPa(N/mm²) × mm² ÷ 1000 = kN。
*)
FUNCTION FC_DL_CompactionPressureCalc : REAL
VAR_INPUT
    fGreenDensGcm3 : REAL;   (* 压坯密度 [g/cm³] Green compact density *)
    fAppDensGcm3   : REAL;   (* 松装密度 [g/cm³] Apparent density *)
    fMatKMPa       : REAL;   (* 材料压制常数 [MPa] Material compaction constant *)
    fPartAreaMm2   : REAL;   (* 压坯投影面积 [mm²] Compact projected area *)
    fSafetyFactor  : REAL;   (* 压机吨位安全系数 [-] Press tonnage safety factor *)
END_VAR
VAR_OUTPUT
    fRelDensity : REAL;   (* 相对密度（压坯/松装） [-] Relative density *)
    fPressMPa   : REAL;   (* 单位压制压力 [MPa] Compaction pressure *)
    fTonnageKN  : REAL;   (* 压机吨位需求 [kN] Required press tonnage *)
    xValid      : BOOL;   (* 计算有效性标志 [-] Calculation valid flag *)
END_VAR
VAR CONSTANT
    DL_EPS      : REAL := 1.0E-9;   (* 除零判定容差 [无量纲] Divide-by-zero tolerance *)
    DL_N_PER_KN : REAL := 1000.0;   (* 牛转千牛系数 [N/kN] Newtons per kilonewton *)
    DL_ONE      : REAL := 1.0;      (* 单位常数 [-] Unity constant *)
    DL_ZERO     : REAL := 0.0;      (* 零常量 [无量纲] Zero constant *)
END_VAR
(* 出口预置：四出口统一预置 *)
fRelDensity := 0.0; fPressMPa := 0.0; fTonnageKN := 0.0; xValid := FALSE;
(* 非有限拦截：自反判 NaN，自身差值判 Inf *)
IF (fGreenDensGcm3 <> fGreenDensGcm3) OR ((fGreenDensGcm3 - fGreenDensGcm3) <> 0.0)
   OR (fAppDensGcm3 <> fAppDensGcm3) OR ((fAppDensGcm3 - fAppDensGcm3) <> 0.0)
   OR (fMatKMPa <> fMatKMPa) OR ((fMatKMPa - fMatKMPa) <> 0.0)
   OR (fPartAreaMm2 <> fPartAreaMm2) OR ((fPartAreaMm2 - fPartAreaMm2) <> 0.0)
   OR (fSafetyFactor <> fSafetyFactor) OR ((fSafetyFactor - fSafetyFactor) <> 0.0) THEN
    FC_DL_CompactionPressureCalc := -1.0;  (* 哨兵 -1：输入非有限 / Sentinel -1 non-finite *)
    RETURN;
END_IF
(* 组态域闸：松装密度为除子，材料常数/面积/安全系数须为正 *)
IF (fAppDensGcm3 <= DL_EPS) OR (fMatKMPa <= DL_ZERO) OR (fPartAreaMm2 <= DL_EPS)
   OR (fSafetyFactor <= DL_ZERO) OR (fGreenDensGcm3 < DL_ZERO) THEN
    FC_DL_CompactionPressureCalc := -1.0;  (* 哨兵 -1：组态非法 / Sentinel -1 bad config *)
    RETURN;
END_IF
(* 相对密度：rho_rel = 压坯密度 / 松装密度，分母已过域闸 *)
fRelDensity := fGreenDensGcm3 / fAppDensGcm3;
IF fRelDensity <= DL_ONE THEN
    xValid := TRUE;                       (* 合法空工况：未致密化，无压制压力 *)
    FC_DL_CompactionPressureCalc := DL_ZERO;
    RETURN;
END_IF
(* 单位压制压力：p = K·(rho_rel - 1) [MPa] *)
fPressMPa := fMatKMPa * (fRelDensity - DL_ONE);
(* 压机吨位需求：p(N/mm²) × A(mm²) = N，除 1000 得 kN，再乘安全系数 *)
fTonnageKN := fPressMPa * fPartAreaMm2 / DL_N_PER_KN * fSafetyFactor;
xValid := TRUE;                           (* 链路有效 / Chain valid *)
FC_DL_CompactionPressureCalc := fPressMPa;  (* 返回压制压力 [MPa] / Return compaction pressure *)
END_FUNCTION
